(* IEC 61131-3 sources: Caravan/Archiv/12-04-19/Stations/MachineControl/MachineControl/Class/SafetyManager (part 2) *)

	state := READY;

//=================================================================================================
#ifdef VM_CLASS_TIME_MEASUREMENT
	StopTimeMeasurement(VARANTIME_CY);
#endif
//=================================================================================================

END_FUNCTION

FUNCTION SafetyManager::AddModule
	VAR_INPUT
		pPara 	: ^CmdStruct;
	END_VAR
	VAR_OUTPUT
		retcode 	: BOOL;
	END_VAR
  VAR
  	ModuleType : t_e_ModuleType;
  END_VAR

  retcode := FALSE;

  ModuleType := pPara^.aPara[0]$t_e_ModuleType;

  // we differ between real safety components and managing components
  case ModuleType of
    _CSCP01x,
    _CSDI16x,
    _CSTO08x,
    _SCP010,
    _SCP011,
    _SCP111,
    _MS011,
    _MS012,
    _SDD1300,
    _SDD1400,
    _SDD1500,
    _SDD1600:
        retcode := AddSafetyModule(ModuleType, pPara^.aPara[1]$pVirtualBase);

        if IsFSoEModule(ModuleType) then
          // allocate memory for the temporary cyclic send buffer
          sUdpVars.pTempSendBufferCy$pVoid := To_StdLib.Malloc(size:=sizeof(t_UdpPacket));

          if sUdpVars.pTempSendBufferCy then
            _memset(dest:=sUdpVars.pTempSendBufferCy, usByte:=0, cntr:=sizeof(t_UdpPacket));
          else
            SetError(bError:=TRUE, ErrorMessage:=_NO_MEMORY_SENDBUFFER_UDP_ERROR, dError:=0);
            LogError("@ZZZZ (SafetyManager::AddModule) Failed to allocate memory for udp send buffer");
          end_if;

          // allocate memory for the temporary irq send buffer
          sUdpVars.pTempSendBufferIRQ$pVoid := To_StdLib.Malloc(size:=sizeof(t_UdpPacket));

          if sUdpVars.pTempSendBufferIRQ then
            _memset(dest:=sUdpVars.pTempSendBufferIRQ, usByte:=0, cntr:=sizeof(t_UdpPacket));
          else
            SetError(bError:=TRUE, ErrorMessage:=_NO_MEMORY_SENDBUFFER_UDP_ERROR, dError:=0);
            LogError("@ZZZZ (SafetyManager::AddModule) Failed to allocate memory for udp send buffer");
          end_if;

          sUdpVars.paConnectionsToProducers$pVoid := To_StdLib.Malloc(size:=sizeof(t_aUdpConnections));

          if sUdpVars.paConnectionsToProducers then
            _memset(dest:=sUdpVars.paConnectionsToProducers, usByte:=0, cntr:=sizeof(t_aUdpConnections));
          else
            SetError(bError:=TRUE, ErrorMessage:=_NO_MEMORY_CONNECTION_BUFFER_UDP_ERROR, dError:=0);
            LogError("@ZZZZ (SafetyManager::AddModule) Failed to allocate memory for udp receive buffer");
          end_if;

          sUdpVars.paConnectionsToConsumers$pVoid := To_StdLib.Malloc(size:=sizeof(t_aUdpConnections));

          if sUdpVars.paConnectionsToConsumers then
            _memset(dest:=sUdpVars.paConnectionsToConsumers, usByte:=0, cntr:=sizeof(t_aUdpConnections));
          else
            SetError(bError:=TRUE, ErrorMessage:=_NO_MEMORY_CONNECTION_BUFFER_UDP_ERROR, dError:=0);
            LogError("@ZZZZ (SafetyManager::AddModule) Failed to allocate memory for udp receive buffer");
          end_if;
        end_if;

    _VBC021Master,
    _VBC021Slave, // (is limited to 1 per system, because the system can't sync to different systems at the same time)
    _VMC052,
    _VaranManager4VMC, // VaranManager (VMC052 counterpart is also limited to 1 per system, because the system can't sync to different systems at the same time)
    _GenericTimeSyncMaster,
    _GenericTimeSyncSlave:
        retcode := AddManagingModule(ModuleType, pPara^.aPara[1]$pVirtualBase, pPara^.aPara[2]$^USINT);
  else
    // invalid module type
    ClassState := -7;
    LogError("@ZZZZ (SafetyManager::AddModule) Invalid ModuleType");
  end_case;

  if retcode then
    LoginCnt += 1;
  end_if;

END_FUNCTION

FUNCTION SafetyManager::AddSafetyModule
	VAR_INPUT
		ModuleType 	: t_e_ModuleType;
		pThis 	: pVirtualBase;
	END_VAR
	VAR_OUTPUT
		retcode 	: BOOL;
	END_VAR
  VAR
  	pHelpSafety : ^t_SafetyComponent;
  END_VAR

  if pFirstSafetyComponent = NIL then
    pFirstSafetyComponent$pVoid := To_StdLib.Malloc(size:=sizeof(t_SafetyComponent));
    pHelpSafety := pFirstSafetyComponent;
  else
    pHelpSafety := pFirstSafetyComponent;
    while pHelpSafety^.pNext <> NIL do
      pHelpSafety := pHelpSafety^.pNext;
    end_while;
    pHelpSafety^.pNext$pVoid := To_StdLib.Malloc(size:=sizeof(t_SafetyComponent));
    pHelpSafety := pHelpSafety^.pNext;
  end_if;

  if pHelpSafety <> NIL then
    _memset(dest:=pHelpSafety, usByte:=0, cntr:=sizeof(t_SafetyComponent));
    pHelpSafety^.ModuleType   := ModuleType;
    pHelpSafety^.pThis        := pThis;

//    pHelpSafety^.pNext        := NIL;  // not necessary because of memset

    case ModuleType of
//**********************************************************************************************************************************************************
      _CSCP01x,
      _SCP010,
      _SCP011,
      _SCP111,
      _SDD1300,
      _SDD1400,
      _SDD1500,
      _SDD1600:
        LocalCPUNo += 1;

//**********************************************************************************************************************************************************
      _CSDI16x,
      _MS011,
      _MS012:
        pHelpSafety^.InfoBits.OnlyInputs := TRUE;
//**********************************************************************************************************************************************************
    end_case;

    us_SafetyModuleNo += 1;

    retcode := TRUE;
  else
    ClassState := -1;

    retcode := FALSE;
  end_if;

END_FUNCTION

FUNCTION SafetyManager::AddManagingModule
	VAR_INPUT
		ModuleType 	: t_e_ModuleType;
		pThis 	: pVirtualBase;
		pObjectPath 	: ^USINT;
	END_VAR
	VAR_OUTPUT
		retcode 	: BOOL;
	END_VAR
  VAR
  	pHelpManaging : ^t_ManagingComponent;
    pMyPath : ^USINT;
  END_VAR

  if pFirstManagingInterfaceComponent = NIL then
    pFirstManagingInterfaceComponent$pVoid := To_StdLib.Malloc(size:=sizeof(t_ManagingComponent));
    pHelpManaging := pFirstManagingInterfaceComponent;
  else
    pHelpManaging := pFirstManagingInterfaceComponent;
    while pHelpManaging^.pNext <> NIL do
      pHelpManaging := pHelpManaging^.pNext;
    end_while;
    pHelpManaging^.pNext$pVoid := To_StdLib.Malloc(size:=sizeof(t_ManagingComponent));
    pHelpManaging := pHelpManaging^.pNext;
  end_if;

  if pHelpManaging <> NIL then
    _memset(dest:=pHelpManaging, usByte:=0, cntr:=sizeof(t_ManagingComponent));
    pHelpManaging^.ModuleType     := ModuleType;
    pHelpManaging^.pThis          := pThis;
    pHelpManaging^.DomainNr       := 16#FF;

    if pObjectPath then
      pMyPath$^void := To_StdLib.Malloc(size:=pObjectPath^ + 2);

      // convert 1 byte length info into 2 byte length info
      if pMyPath then
        pMyPath^$UINT := pObjectPath^$USINT;
        To_StdLib.MemCpy(dest:=pMyPath + 2, source:=pObjectPath + 1, size:=pObjectPath^);
      end_if;
    end_if;

    pHelpManaging^.pModulePath := pMyPath;

  //pHelpManaging^.pNext          := NIL;  // not necessary because of memset

    retcode := TRUE;
  else
    ClassState := -1;

    retcode := FALSE;
  end_if;

END_FUNCTION

FUNCTION SafetyManager::AddSafetyNbr
	VAR_INPUT
		pThis 	: pVirtualBase;
		ud_SafetyNbr 	: UDINT;
		FirmwareVersion 	: HDINT;
		FPGAVersion 	: HSINT;
		PathLen 	: USINT;
		pPath 	: ^USINT;
	END_VAR
	VAR_OUTPUT
		retcode 	: BOOL;
	END_VAR
  VAR
  	pHelpSafety : ^t_SafetyComponent;
  END_VAR

  retcode := FALSE;

  if pFirstSafetyComponent then
    pHelpSafety := pFirstSafetyComponent;
    while pHelpSafety do
      if pHelpSafety^.pThis = pThis then
        pHelpSafety^.SafetyNbr    := ud_SafetyNbr;
        pHelpSafety^.FW_Version   := FirmwareVersion;
        pHelpSafety^.FPGA_Version := FPGAVersion;
        pHelpSafety^.PathLen      := PathLen;
        pHelpSafety^.pPath        := pPath;

        // look for local safety CPU
        if b_CheckSafetyTopology then
          if (PathLen > 2) & (((pPath+2)^ = HWT_ESCAPE_CDIAS) | ((pPath+2)^ = HWT_ESCAPE_SDIAS)) then
            b_CheckSafetyTopology := FALSE; // Safety-CPU is local -> no problem
          end_if;
        end_if;

        retcode := TRUE;
        return;
      end_if;

      pHelpSafety := pHelpSafety^.pNext;
    end_while;
  end_if;

END_FUNCTION

FUNCTION SafetyManager::GetModuleTypeNo
	VAR_INPUT
		ModuleType 	: t_e_ModuleType;
	END_VAR
	VAR_OUTPUT
		ModuleNo 	: DINT;
	END_VAR
  VAR
  	pHelpSafety   : ^t_SafetyComponent;
    pHelpManaging : ^t_ManagingComponent;
  END_VAR

  ModuleNo := 0;

  if pFirstSafetyComponent then
    pHelpSafety := pFirstSafetyComponent;
    while pHelpSafety do
      if pHelpSafety^.ModuleType = ModuleType then
        ModuleNo += 1;
      end_if;

      pHelpSafety := pHelpSafety^.pNext;
    end_while;
  end_if;

  if pFirstManagingInterfaceComponent then
    pHelpManaging := pFirstManagingInterfaceComponent;
    while pHelpManaging do
      if pHelpManaging^.ModuleType = ModuleType then
        ModuleNo += 1;
      end_if;

      pHelpManaging := pHelpManaging^.pNext;
    end_while;
  end_if;

END_FUNCTION

FUNCTION SafetyManager::NewTimeSyncPossible
	VAR_OUTPUT
		retcode 	: BOOL;
	END_VAR
  VAR
  	pHelpSafety   : ^t_SafetyComponent;
  END_VAR

  // if there is FSoE in the project => no timesync
  if b_GotFSoEModules then
    retcode := FALSE;
    return;
  end_if;

  // default is: we can => check if there is any module with too old firmware or fpga
  retcode := TRUE;

  if pFirstSafetyComponent then
    pHelpSafety := pFirstSafetyComponent;
    while pHelpSafety do

      // check all modules for correct versions
      if ((pHelpSafety^.ModuleType = _CSCP01x) & (   (pHelpSafety^.FPGA_Version    < 16#14)     // if its a CSCP and the FPGA Version is lower than 1.4
                                                   | (pHelpSafety^.FW_Version$UINT < 100)) &    // or the firmware version is lower than 100
                                                      pHelpSafety^.SafetyNbr)                   // only if there is a safety number available (maybe the module is optional and not available)
      |  (pHelpSafety^.NewConfigType = ConfigState_Old) then                                    // or the module has an old config type

        retcode := FALSE;
      end_if;

      pHelpSafety := pHelpSafety^.pNext;
    end_while;
  end_if;

END_FUNCTION

FUNCTION SafetyManager::SetNewSyncMode
	VAR_INPUT
		b_NewMode 	: BOOL;
	END_VAR
  VAR
		MyPara 	  : CmdStruct;
		MyResult	: results;
  END_VAR

  b_NewSyncMode := b_NewMode;

  MyPara.uiCmd := CMD_SM_SET_NEW_SYNC_MODE;
  MyPara.aPara[0] := b_NewSyncMode;
  TellAllSafetyModules(#MyPara, #MyResult);

END_FUNCTION

FUNCTION SafetyManager::TellAllSafetyModules
	VAR_INPUT
		pPara 	: ^CmdStruct;
		pResult 	: ^results;
	END_VAR
  VAR
  	pHelpSafety : ^t_SafetyComponent;
  END_VAR

  if pFirstSafetyComponent then
    pHelpSafety := pFirstSafetyComponent;
    while pHelpSafety do
      // call the newinst with the given parameters
      pHelpSafety^.pThis^.NewInst(pPara, pResult);

      pHelpSafety := pHelpSafety^.pNext;
    end_while;
  end_if;

END_FUNCTION

FUNCTION SafetyManager::StartTimeSync

  if pFirstTimeSyncElement then
    pActTimeSyncElement := pFirstTimeSyncElement;

    // send the token to the right module
    GiveTokenToNextModule();

    // remember the start time for calculating the time of a complete synchronisation
    TimeSyncCycleStart := ops.tAbsolute;
  end_if;

END_FUNCTION

FUNCTION SafetyManager::NextTimeSyncModule

  pActTimeSyncElement := pActTimeSyncElement^.pNext;

  // must be done after selecting the new element
  if GiveTokenToNextModule() then
    // we're finished with our synchronisation cycle and just started a new one (must be done after selecting the new element)
    if IsTimeSyncMaster then
      SyncDuration := ops.tAbsolute - TimeSyncCycleStart;
      if SyncDuration > MaxSyncDuration then
        MaxSyncDuration := SyncDuration;
      end_if;
      if SyncDuration < MinSyncDuration then
        MinSyncDuration := SyncDuration;
      end_if;

      // if a cycle has been finished => reset the timeout counter
      SyncTimeoutCounter := 0;

      // remember the start time for calculating the time of a complete synchronisation
      TimeSyncCycleStart := ops.tAbsolute;
    end_if;
  end_if;

END_FUNCTION

FUNCTION SafetyManager::GiveTokenToNextModule
	VAR_OUTPUT
		RestartCycle 	: BOOL;
	END_VAR
  VAR
		MyPara 	  : CmdStruct;
		MyResult	: results;
    pTemp : ^t_TimeSyncElement;
  END_VAR

  if pActTimeSyncElement = pFirstTimeSyncElement then
    RestartCycle := TRUE;
  else
    RestartCycle := FALSE;
  end_if;

  // check if we have to skip something (missing optional modules)
  if TimeSyncModuleAvailable(pActTimeSyncElement) = FALSE then
    // save the actual position
    pTemp := pActTimeSyncElement;

    // if it's a missing optional module
    while (TimeSyncModuleAvailable(pActTimeSyncElement) = FALSE) do
      // skip it
      pActTimeSyncElement := pActTimeSyncElement^.pNext;

      // if we jumped on the first, we have to restart the cycle (time measurement and timeout surveillance)
      if pActTimeSyncElement = pFirstTimeSyncElement then
        RestartCycle := TRUE;
      end_if;

      // if we're at the start of the rotation => stop rotating and print error message
      if pActTimeSyncElement = pTemp then
        bd_LogRtMessagesInCy.TooManyOptionalMissing := TRUE;
        ClassState := -12;
        exit;
      end_if;
    end_while;
  end_if;

  // check if we have to skip something
  if pActTimeSyncElement^.InfoBits.IsInterfaceDomain then
    // save the actual position
    pTemp := pActTimeSyncElement;

    // if it's an interface managing module and it's not synchron, skip it (there has to be also a Safety CPU in the system, therefore we don't ask for it
    while pActTimeSyncElement^.InfoBits.IsInterfaceDomain & (pActTimeSyncElement^.pManaging^.InfoBits.IsSynchron = FALSE) do
      // skip it
      pActTimeSyncElement := pActTimeSyncElement^.pNext;

      // if we jumped on the first, we have to restart the cycle (time measurement and timeout surveillance)
      if pActTimeSyncElement = pFirstTimeSyncElement then
        RestartCycle := TRUE;
      end_if;

      // if we're at the start of the rotation => stop rotating and print error message
      if pActTimeSyncElement = pTemp then
        bd_LogRtMessagesInCy.InvalidIFConfiguration := TRUE;
        ClassState := -12;
        exit;
      end_if;
    end_while;
  end_if;

  if pActTimeSyncElement^.InfoBits.IsConnectionToMaster then
    // don't check for sync timeout if we're not the master
    b_CheckTimeSyncTimeout := FALSE;
  else
    b_CheckTimeSyncTimeout := TRUE;
  end_if;

  // if it's a managing module and not the connection to the master, we give the token to a slave => remember it
  if pActTimeSyncElement^.InfoBits.IsManagingModule & (pActTimeSyncElement^.InfoBits.IsConnectionToMaster = FALSE) then
    b_SlaveSyncActive := TRUE;
  end_if;

  // tell the next module, to start the time synchronisation
  MyPara.uiCmd := CMD_SM_START_TIME_SYNC;
  pActTimeSyncElement^.pThis^.NewInst(#MyPara, #MyResult);

  LastTimeSyncThis := pActTimeSyncElement^.pThis;
  TimeSyncTimeStamp := ops.tAbsolute;

END_FUNCTION

FUNCTION SafetyManager::TellAllInterfaceManagingModules
	VAR_INPUT
		pPara 	: ^CmdStruct;
		pResult 	: ^results;
		OverrideSync 	: BOOL;(* := FALSE *)
	END_VAR
  VAR
  	pHelpManaging : ^t_ManagingComponent;
  END_VAR

  if pFirstManagingInterfaceComponent then
    pHelpManaging := pFirstManagingInterfaceComponent;
    while pHelpManaging do
      // call the newinst with the given parameters
      if pHelpManaging^.InfoBits.IsSynchron | OverrideSync then
        pHelpManaging^.pThis^.NewInst(pPara, pResult);
      end_if;

      pHelpManaging := pHelpManaging^.pNext;
    end_while;
  end_if;

END_FUNCTION

FUNCTION SafetyManager::SafetyManager
	VAR_OUTPUT
		ret_code 	: ConfStates;
	END_VAR
  VAR
    sd_retval : DINT;
  END_VAR

  //get interface for hardwaretree functions
  if ( OS_CILGET(INTERFACE_HARDWARETREE, #pHardwareTree)) then
    pHardwareTree := NIL;

    // logging can be used here already because the constructor of the base has been called before to initialize the log-interface-pointer
    LogError("@ZZZZ (SafetyManager::SafetyManager) Hardwaretree-Interface not found. A newer OS is required for Safety-Modules");
  end_if;

  pTempMemCy := To_StdLib.Malloc(size:=SIZE_TEMP_MEMORY);
  if pTempMemCy then
    ud_SizeTempMemCy := SIZE_TEMP_MEMORY;
  else
    LogError("@ZZZZ (SafetyManager::SafetyManager) Allocate temporary Memory failed");
  end_if;

  b_QuitErrorAvailable := FALSE;

  sd_retval := OS_CILGet(INTERFACE_SAFETY_DLL, #pSafetyDll)$DINT;

  if sd_retval then
    // normal case => no dll available
//    LogValue("@ZZZZ (SafetyManager::SafetyManager) Failed to get interface to safety DLL with ErrorCode 0x{0}", Value:=sd_retval$UDINT);
  elsif pSafetyDll^.version >= 5 then
//    LogValue("@ZZZZ (SafetyManager::SafetyManager) Safety DLL with Version 0x{0} loaded. QuitError via Application available!", Value:=pSafetyDll^.version);

    b_QuitErrorAvailable := TRUE;
  end_if;

  // as long there is no Safety-CPU on local CDIAS or SDIAS, we need to check for "unalowed" safety communication over VARAN.
  b_CheckSafetyTopology := TRUE;
  OS_CILGet( INTERFACE_VARANMANAGER, #pVaran );

	ret_code := C_OK;

END_FUNCTION

FUNCTION SafetyManager::AllManagingNodesSynchron
	VAR_OUTPUT
		AllReady 	: BOOL;
	END_VAR
  VAR
  	pHelpManaging : ^t_ManagingComponent;
		MyPara 	  : CmdStruct;
		MyResult	: results;
  END_VAR

  AllReady := TRUE;

  // check if any of the managing interface modules is not synchron
  if pFirstManagingInterfaceComponent then
    MyPara.uiCmd := CMD_SM_SYNC_CHECK;

    pHelpManaging := pFirstManagingInterfaceComponent;
    while pHelpManaging do
      // if any managing component isn't synchron => stop searching
      if pHelpManaging^.pThis^.NewInst(#MyPara, #MyResult) = ERROR then
        if (pHelpManaging^.InfoBits.IsOptional = TRUE) then
          if ((SafetyDomainTimeout & ((ops.tAbsolute - SynchroTimeout) > SafetyDomainTimeout))) then
            // we give up waiting => timeout exceeded
            b_SyncTimeoutExceeded := TRUE;
            // if it's the last managing module, then it's our connection to the master module
            if (IsTimeSyncMaster = 0) & pHelpManaging^.InfoBits.IsConnectionToMaster then
              // we have to be our own master now
              IsTimeSyncMaster := 1;
            end_if;
          else
            AllReady := FALSE;
          end_if;
        else
          AllReady := FALSE;
        end_if;

        // return; don't give up here => we have to check it for all domains, this one may be an optional interface frame domain
        pHelpManaging^.InfoBits.IsSynchron := FALSE;
      else
        pHelpManaging^.InfoBits.IsSynchron := TRUE;
      end_if;

      pHelpManaging := pHelpManaging^.pNext;
    end_while;
  end_if;

END_FUNCTION

FUNCTION SafetyManager::GetMasterConnection
  VAR_OUTPUT
    pMasterConn : ^t_ManagingComponent;
  END_VAR
  VAR
    pHelpManaging : ^t_ManagingComponent;
  END_VAR

  pMasterConn := NIL;

  if pFirstManagingInterfaceComponent then
    pHelpManaging := pFirstManagingInterfaceComponent;
    while pHelpManaging do
      if (pHelpManaging^.ModuleType = _VBC021Slave) | (pHelpManaging^.ModuleType = _VaranManager4VMC) | (pHelpManaging^.ModuleType = _GenericTimeSyncSlave) then
        pMasterConn := pHelpManaging;
        pMasterConn^.InfoBits.IsConnectionToMaster := TRUE;
        // if it's not the last in the list => we have to put it in the last place for easier timesync handling (last managing module to handle is the connection back to the master)
        if pMasterConn^.pNext then
          // if it's the first one
          if pMasterConn = pFirstManagingInterfaceComponent then
            pHelpManaging := pFirstManagingInterfaceComponent;
            while pHelpManaging^.pNext do
              pHelpManaging := pHelpManaging^.pNext;
            end_while;
            pFirstManagingInterfaceComponent := pFirstManagingInterfaceComponent^.pNext;
            pHelpManaging^.pNext := pMasterConn;
            pMasterConn^.pNext := NIL;
          else
            // if it's one in the middle
            pHelpManaging := pFirstManagingInterfaceComponent;
            while pHelpManaging^.pNext do
              if pHelpManaging^.pNext = pMasterConn then
                pHelpManaging^.pNext := pMasterConn^.pNext;
              end_if;

              pHelpManaging := pHelpManaging^.pNext;
            end_while;
            pHelpManaging^.pNext := pMasterConn;
            pMasterConn^.pNext := NIL;
          end_if;
        end_if;
        return;
      end_if;

      pHelpManaging := pHelpManaging^.pNext;
    end_while;
  end_if;

END_FUNCTION

FUNCTION SafetyManager::AddConfiguration
	VAR_INPUT
		Length 	: UINT;
		pData 	: ^void;
		IsFSoEConfig 	: BOOL;
	END_VAR
	VAR_OUTPUT
		retcode 	: DINT;
	END_VAR
  VAR
    pHelpCfg          : ^t_CfgListElem;
    pHelpModule       : ^t_ModuleListElem;
    pHelpPdo          : ^t_PdoListElem;
    pHelpSlave        : ^t_SlaveListElem;
    pHelpConnection   : ^t_FSoEConnectionDetails;
    pDataHelp         : ^void;
    i                 : UDINT;
    TmpPathLen        : UINT;
    TempCfgNo         : USINT;
    TempConnectionNo  : UINT;
  END_VAR

(*
    Memory structure:
      4 Byte: SafetyNumber of CPU (is already there from initialisation in CSCP011_IM::InitSafeModule)
      1 Byte: Number of module configurations which are following
      for every module configuration (first is always the CPU itself)
        1 Byte: Info
        4 Byte: Interface Frame Source SafetyNumber (0 if it is no source for interface frames)
        4 Byte: Interface Frame CRC
        1 Byte: Number of destination inferface frame CRCs
        x Byte: Destination interface frame CRCs (number * sizeof(HDINT)
        2 Byte: Length of hardware path
        x Byte (depending on length in the 2 byte before): Hardwarepath
        2 Byte: Length of compressed hardware path
        x Byte (depending on length in the 2 byte before): Compressed Hardwarepath
        1 Byte: PDO out length for this module
      1 Byte: Number of pdo configurations which are following
      for every PDO configuration
        1 Byte: PDO length
        1 Byte: Interface frame info
        4 Byte: Interface CRC
        2 Byte: Length of source hardware path
        x Byte (depending on length in the 2 byte before): Hardwarepath of source
        2 Byte: Length of destination hardware path
        x Byte (depending on length in the 2 byte before): Hardwarepath of destination
      1 Byte: Number of slave configurations which are following
      for every slave configuration
        1 Byte: Info
        4 Byte: InterfaceCRC
        2 Byte: Length of hardware path
        x Byte (depending on length in the 2 byte before): Hardwarepath
        2 Byte: Length of compressed hardware path
        x Byte (depending on length in the 2 byte before): Compressed Hardwarepath

      if IsFSoEConfig = TRUE
      2 Byte: Number of connection infos which are following
      for every FSoE connection info
        2 Byte: ConnectionID
        1 Byte: ConnectionState
        1 Byte: Flags // Actually, type is 4 bytes in size but for compatibility reasons it is still used as 1 byte. As a result, bits 9-32 are currently not used.
        4 Byte: Master safety number

only if feature available:
        2 Byte: Transmission time in ms

        2 Byte: Offset where to read from master
        2 Byte: Size of data to read from master (and write to slave)
        2 Byte: Offset where to write to master
        2 Byte: Size of data to write to master (and read from slave)
        2 Byte: SlaveAddress
        2 Byte: Length of slave hardware path
        x Byte (depending on length in the 2 byte before): Slave hardware path
        2 Byte: Length of compressed slave hardware path
        x Byte (depending on length in the 2 byte before): Compressed slave hardware path
        2 Byte: Offset where to read from slave
        2 Byte: Offset where to write to slave

*)

  // check if the configuration is valid (pData <> NIL) & (Length must be at least 4 byte for SafetyNbr + 1 byte module cfg number + 1 byte pdo cfg number + 1 byte slave cfc number)
  if pData & (Length >= 7)  then

    retcode := 0;

    // first we have to allocate some memory for the configuration
    if pConfigs = NIL then
      pConfigs$pVoid := To_StdLib.Malloc(size:=sizeof(t_CfgListElem));
      pHelpCfg := pConfigs;
    else
      pHelpCfg := pConfigs;
      while pHelpCfg^.pNext <> NIL do
        //if searched path is found, we already got this module in our list
        if pHelpCfg^.SafetyNbr = pData^$HDINT then
          // already in buffer => leave function
          return;
        else
          pHelpCfg := pHelpCfg^.pNext;
        end_if;
      end_while;

      //if searched path is found, we already got this module in our list
      if pHelpCfg^.SafetyNbr = pData^$HDINT then
        // already in buffer => leave function
        return;
      end_if;

      pHelpCfg^.pNext$pvoid := To_StdLib.Malloc(size:=sizeof(t_CfgListElem));
      pHelpCfg := pHelpCfg^.pNext;
    end_if;

    // if we have memory for the configuration => we add the data to the new element
    if pHelpCfg <> NIL then
      pDataHelp := pData;

      // set the next pointer to NIL
      pHelpCfg^.pNext := NIL;

      // safety number of the safety cpu
      pHelpCfg^.SafetyNbr := pDataHelp^$HDINT;
      pDataHelp += sizeof(HDINT);

      // number of module configurations which follow now
      TempCfgNo := pDataHelp^$USINT;
      pDataHelp += sizeof(USINT);

      pHelpCfg^.pFirstModuleCfg := NIL;

      // module configurations
      if TempCfgNo then
        for i := 0 to (TempCfgNo-1) do
          if pHelpCfg^.pFirstModuleCfg = NIL then
            pHelpCfg^.pFirstModuleCfg$pVoid := To_StdLib.Malloc(size:=sizeof(t_ModuleListElem));
            pHelpModule := pHelpCfg^.pFirstModuleCfg;
          else
            pHelpModule^.pNext$pvoid := To_StdLib.Malloc(size:=sizeof(t_ModuleListElem));
            pHelpModule := pHelpModule^.pNext;
          end_if;

          if pHelpModule then
            // initialize the pointers with NIL in case one of the mallocs fails
            pHelpModule^.ModuleInfo.pDestCRCs   := NIL;
            pHelpModule^.ModuleInfo.pPath       := NIL;
            pHelpModule^.ModuleInfo.pCompPath   := NIL;
            pHelpModule^.pNext                  := NIL;

            // info
            pHelpModule^.ModuleInfo.Info := pDataHelp^$BSINT;
            pDataHelp += sizeof(BSINT);

            // safety number of interface frame source
            pHelpModule^.ModuleInfo.SafetyNbr := pDataHelp^$HDINT;
            pDataHelp += sizeof(HDINT);

            // interface CRC of interface frame
            pHelpModule^.ModuleInfo.InterfaceCRC := pDataHelp^$HDINT;
            pDataHelp += sizeof(HDINT);

            if pHelpModule^.ModuleInfo.InterfaceCRC then
              // someone might connect to us via udp because we supply an interface frame
              sUdpVars.UdpInit.ProvidesIF := TRUE;
            end_if;

            // interface frame destination CRCs
            if pHelpModule^.ModuleInfo.Info.IsInterfaceDest then
              // number of CRCs
              TmpPathLen := pDataHelp^$USINT; // save some time with this local variable
              pHelpModule^.ModuleInfo.DestCRCNo := TmpPathLen$USINT;
              pDataHelp += sizeof(USINT);

              // allocate memory for the module path
              pHelpModule^.ModuleInfo.pDestCRCs$pVoid := To_StdLib.Malloc(size:=TmpPathLen * sizeof(HDINT));
              if pHelpModule^.ModuleInfo.pDestCRCs = NIL then
                ClassState := -1;
                retcode := -2;
                return;
              end_if;

              // save CRCs
              _memcpy(ptr1:=pHelpModule^.ModuleInfo.pDestCRCs, ptr2:=pDataHelp, cntr:=TmpPathLen * sizeof(HDINT));
              pDataHelp += TmpPathLen * sizeof(HDINT);
            else
              pHelpModule^.ModuleInfo.DestCRCNo := 0;
              pHelpModule^.ModuleInfo.pDestCRCs := NIL;
            end_if;

            // length of hardwarepath
            TmpPathLen := pDataHelp^$UINT; // save some time with this local variable
            pHelpModule^.ModuleInfo.PathLen := TmpPathLen;
            pDataHelp += sizeof(UINT);

            // allocate memory for the module path
            pHelpModule^.ModuleInfo.pPath$pVoid := To_StdLib.Malloc(size:=TmpPathLen);
            if pHelpModule^.ModuleInfo.pPath = NIL then
              ClassState := -1;
              retcode := -2;
              return;
            end_if;

            // save hardwarepath
            _memcpy(ptr1:=pHelpModule^.ModuleInfo.pPath, ptr2:=pDataHelp, cntr:=TmpPathLen);
            pDataHelp += TmpPathLen;

            // length of hardwarepath
            TmpPathLen := pDataHelp^$UINT; // save some time with this local variable
            pHelpModule^.ModuleInfo.CompPathLen := TmpPathLen;
            pDataHelp += sizeof(UINT);

            // allocate memory for the module path
            pHelpModule^.ModuleInfo.pCompPath$pVoid := To_StdLib.Malloc(size:=TmpPathLen);
            if pHelpModule^.ModuleInfo.pCompPath = NIL then
              ClassState := -1;
              retcode := -2;
              return;
            end_if;

            // save compressed hardwarepath
            _memcpy(ptr1:=pHelpModule^.ModuleInfo.pCompPath, ptr2:=pDataHelp, cntr:=TmpPathLen);
            pDataHelp += TmpPathLen;

            // PDO out length for this module (to assign the length to the pdo configurations)
            pHelpModule^.ModuleInfo.PdoOutLen := pDataHelp^$USINT;
            pDataHelp += sizeof(USINT);
          else
            ClassState := -1;
            retcode := -2;
            return;
          end_if;
        end_for;
      end_if;

      // number of Pdo configurations which follow now
      TempCfgNo := pDataHelp^$USINT;
      pDataHelp += sizeof(USINT);

      pHelpCfg^.pFirstPdoCfg := NIL;

      // Pdo configurations
      if TempCfgNo then
        for i := 0 to (TempCfgNo-1) do
          if pHelpCfg^.pFirstPdoCfg = NIL then
            pHelpCfg^.pFirstPdoCfg$pVoid := To_StdLib.Malloc(size:=sizeof(t_PdoListElem));
            pHelpPdo := pHelpCfg^.pFirstPdoCfg;
          else
            pHelpPdo^.pNext$pvoid := To_StdLib.Malloc(size:=sizeof(t_PdoListElem));
            pHelpPdo := pHelpPdo^.pNext;
          end_if;

          if pHelpPdo then
            // initialize the pointers with NIL in case one of the mallocs fails
            pHelpPdo^.PdoInfo.pSourcePath     := NIL;
            pHelpPdo^.PdoInfo.pDestPath       := NIL;
            pHelpPdo^.pNext                   := NIL;

            // pdo length
            pHelpPdo^.PdoInfo.PdoLen := pDataHelp^$USINT;
            pDataHelp += sizeof(USINT);

            // is it an interface pdo?
            pHelpPdo^.PdoInfo.Info := pDataHelp^$BSINT;
            pDataHelp += sizeof(BSINT);

            // if it is an interface frame, we have to copy the CRC too
            if pHelpPdo^.PdoInfo.Info.IsInterfacePDO then
              // interface CRC
              pHelpPdo^.PdoInfo.InterfaceCRC := pDataHelp^$HDINT;
            else
              pHelpPdo^.PdoInfo.InterfaceCRC := 0;
            end_if;
            pDataHelp += sizeof(HDINT);

            // length of source hardwarepath
            TmpPathLen := pDataHelp^$UINT; // save some time with this local variable
            pHelpPdo^.PdoInfo.SourcePathLen := TmpPathLen;
            pDataHelp += sizeof(UINT);

            // allocate memory for the source module path
            pHelpPdo^.PdoInfo.pSourcePath$pVoid := To_StdLib.Malloc(size:=TmpPathLen);
            if pHelpPdo^.PdoInfo.pSourcePath = NIL then
              ClassState := -1;
              retcode := -2;
              return;
            end_if;

            // save source hardwarepath
            _memcpy(ptr1:=pHelpPdo^.PdoInfo.pSourcePath, ptr2:=pDataHelp, cntr:=TmpPathLen);
            pDataHelp += TmpPathLen;

            // check for an IP Address
            if pHelpPdo^.PdoInfo.Info.SrcPathIsCompressed & (pHelpPdo^.PdoInfo.pSourcePath^$USINT = INTERFACE_IP_MODE) then
              // add the connection (we're consumer and we got the IP address of the producer)
              AddUdpConnection(IP:=(pHelpPdo^.PdoInfo.pSourcePath$^HDINT + 5)^, IFCRC:=(pHelpPdo^.PdoInfo.pSourcePath$^HDINT + 1)^, SafetyNumber:=pHelpCfg^.SafetyNbr, ProducerList:=TRUE);
            end_if;

            // length of destination hardwarepath
            TmpPathLen := pDataHelp^$UINT; // save some time with this local variable
            pHelpPdo^.PdoInfo.DestPathLen := TmpPathLen;
            pDataHelp += sizeof(UINT);

            // allocate memory for the destination module path
            pHelpPdo^.PdoInfo.pDestPath$pVoid := To_StdLib.Malloc(size:=TmpPathLen);
            if pHelpPdo^.PdoInfo.pDestPath = NIL then
              ClassState := -1;
              retcode := -2;
              return;
            end_if;

            // save destination hardwarepath
            _memcpy(ptr1:=pHelpPdo^.PdoInfo.pDestPath, ptr2:=pDataHelp, cntr:=TmpPathLen);
            pDataHelp += TmpPathLen;

            // check if a prior configuration also added this PDO (possible if a CSTO gets PDOs from 2 CSCPs)
            if DoublePDOEntry(pHelpPdo^.PdoInfo, pHelpCfg) then
              // use ID 255 (as kind of invalid) and mark the PDO as double entry (will not be distributed then)
              pHelpPdo^.PdoInfo.PDO_ID := 255;
              pHelpPdo^.PdoInfo.Info.DoublePDOEntry := TRUE;
            else
              // now we give it a priority and increase the number for the next pdo
              pHelpPdo^.PdoInfo.PDO_ID := ActPDO_ID;
              ActPDO_ID += 1;
            end_if;

          else
            ClassState := -1;
            retcode := -2;
            return;
          end_if;
        end_for;
      end_if;

      // number of slave configurations which follow now
      TempCfgNo := pDataHelp^$USINT;
      pDataHelp += sizeof(USINT);

      pHelpCfg^.pFirstSlaveCfg:= NIL;

      // slave configurations
      if TempCfgNo then
        for i := 0 to (TempCfgNo-1) do
          if pHelpCfg^.pFirstSlaveCfg = NIL then
            pHelpCfg^.pFirstSlaveCfg$pVoid := To_StdLib.Malloc(size:=sizeof(t_SlaveListElem));
            pHelpSlave := pHelpCfg^.pFirstSlaveCfg;
          else
            pHelpSlave^.pNext$pvoid := To_StdLib.Malloc(size:=sizeof(t_SlaveListElem));
            pHelpSlave := pHelpSlave^.pNext;
          end_if;

          if pHelpSlave then
            // initialize the pointers with NIL in case one of the mallocs fails
            pHelpSlave^.SlaveInfo.pPath     := NIL;
            pHelpSlave^.SlaveInfo.pCompPath := NIL;
            pHelpSlave^.pNext               := NIL;

            // info
            pHelpSlave^.SlaveInfo.Info := pDataHelp^$BSINT;
            pDataHelp += sizeof(BSINT);

            // InterfaceCRC
            pHelpSlave^.SlaveInfo.InterfaceCRC := pDataHelp^$HDINT;
            pDataHelp += sizeof(HDINT);

            // length of hardwarepath
            TmpPathLen := pDataHelp^$UINT; // save some time with this local variable
            pHelpSlave^.SlaveInfo.PathLen := TmpPathLen;
            pDataHelp += sizeof(UINT);

            // allocate memory for the module path
            pHelpSlave^.SlaveInfo.pPath$pVoid := To_StdLib.Malloc(size:=TmpPathLen);
            if pHelpSlave^.SlaveInfo.pPath = NIL then
              ClassState := -1;
              retcode := -2;
              return;
            end_if;

            // save hardwarepath
            _memcpy(ptr1:=pHelpSlave^.SlaveInfo.pPath, ptr2:=pDataHelp, cntr:=TmpPathLen);
            pDataHelp += TmpPathLen;

            // length of hardwarepath
            TmpPathLen := pDataHelp^$UINT; // save some time with this local variable
            pHelpSlave^.SlaveInfo.CompPathLen := TmpPathLen;
            pDataHelp += sizeof(UINT);

            // allocate memory for the module path
            pHelpSlave^.SlaveInfo.pCompPath$pVoid := To_StdLib.Malloc(size:=TmpPathLen);
            if pHelpSlave^.SlaveInfo.pCompPath = NIL then
              ClassState := -1;
              retcode := -2;
              return;
            end_if;

            // save compressed hardwarepath
            _memcpy(ptr1:=pHelpSlave^.SlaveInfo.pCompPath, ptr2:=pDataHelp, cntr:=TmpPathLen);
            pDataHelp += TmpPathLen;
          else
            ClassState := -1;
            retcode := -2;
            return;
          end_if;
        end_for;
      end_if;

      pHelpCfg^.pFirstFSoEConnection := NIL;

      // check if it's a FSoE Config
      if IsFSoEConfig then
        // number of connection details which follow now
        TempConnectionNo := pDataHelp^$UINT;
        pDataHelp += sizeof(UINT);

        // if we got connections
        if TempConnectionNo then
          for i := 0 to (TempConnectionNo-1) do
            if pHelpCfg^.pFirstFSoEConnection = NIL then
              pHelpCfg^.pFirstFSoEConnection$pVoid := To_StdLib.Malloc(size:=sizeof(t_FSoEConnectionDetails));
              pHelpConnection := pHelpCfg^.pFirstFSoEConnection;
            else
              pHelpConnection^.pNext$pvoid := To_StdLib.Malloc(size:=sizeof(t_FSoEConnectionDetails));
              pHelpConnection := pHelpConnection^.pNext;
            end_if;

            // if we succeeded to allocate memory
            if pHelpConnection then
              // initialize the pointers with NIL in case one of the mallocs fails
              pHelpConnection^.pSlavePath       := NIL;
              pHelpConnection^.pSlavePathComp   := NIL;
              pHelpConnection^.pNext            := NIL;
              pHelpConnection^.pNextSorted      := NIL;

              // connection ID
              pHelpConnection^.ConnectionID := pDataHelp^$UINT;
              pDataHelp += sizeof(UINT);

              // connection state (use our own state internally)
              pHelpConnection^.InternalConnectionState := FCS_RESET;
              pHelpConnection^.ConnectionState := pDataHelp^$t_FSoEConnectionState;

              pDataHelp += sizeof(USINT);

              // flags

              // Actually, type is 4 bytes in size but for compatibility reasons it is still used as 1 byte. As a result, bits 9-32 are currently not used.
              if bdFeatureEnable.FSoEFlags_4ByteSize then
                pHelpConnection^.Flags$t_FSoEFlags := pDataHelp^$t_FSoEFlags;
                pDataHelp += sizeof(t_FSoEFlags);
              else
                pHelpConnection^.Flags$USINT := pDataHelp^$USINT;
                pDataHelp += sizeof(USINT);
              end_if;

              // master safety number
              pHelpConnection^.OwnerSafetyNbr := pDataHelp^$HDINT;
              pDataHelp += sizeof(HDINT);

              // the feature is not available in older safety module classes, so we have to do this for compatibility reasons
              if bdFeatureEnable.TransmissionTimeInConfig then
                // transmission time in ms
                pHelpConnection^.TransmissionTime_ms := pDataHelp^$UINT;
                pDataHelp += sizeof(UINT);
              else
                pHelpConnection^.TransmissionTime_ms := 0;
              end_if;

              // offset where to read from master
              pHelpConnection^.MasterReadOffset := pDataHelp^$UINT;
              pDataHelp += sizeof(UINT);

              // size of data to read from master (and write to slave)
              pHelpConnection^.MasterReadSize := pDataHelp^$UINT;
              pDataHelp += sizeof(UINT);

              // offset where to write to master
              pHelpConnection^.MasterWriteOffset := pDataHelp^$UINT;
              pDataHelp += sizeof(UINT);

              // size of data to write to master (and read from slave)
              pHelpConnection^.MasterWriteSize := pDataHelp^$UINT;
              pDataHelp += sizeof(UINT);

              // slave address
              pHelpConnection^.SlaveAddress := pDataHelp^$UINT;
              pDataHelp += sizeof(UINT);

              // wait for slave addresses if any connection is not initialized
              if (pHelpConnection^.ConnectionState = FCS_NOT_INITIALIZED) & (pHelpConnection^.SlaveAddress = 0) then
                b_AllLocalSlaveAddressesValid := FALSE;
              end_if;

              // length of uncompressed slave hardwarepath
              TmpPathLen := pDataHelp^$UINT; // save some time with this local variable
              pHelpConnection^.SlavePathLen := TmpPathLen;
              pDataHelp += sizeof(UINT);

              if pHelpConnection^.Flags.IsMaster then
                // allocate memory for the module path
                pHelpConnection^.pSlavePath$pVoid := To_StdLib.Malloc(size:=TmpPathLen);
                if pHelpConnection^.pSlavePath = NIL then
                  ClassState := -1;
                  retcode := -2;
                  return;
                end_if;

                // save hardwarepath
                _memcpy(ptr1:=pHelpConnection^.pSlavePath, ptr2:=pDataHelp, cntr:=TmpPathLen);
                pDataHelp += TmpPathLen;
              end_if;

              // length of compressed slave hardwarepath
              TmpPathLen := pDataHelp^$UINT; // save some time with this local variable
              pHelpConnection^.SlavePathCompLen := TmpPathLen;
              pDataHelp += sizeof(UINT);

              if pHelpConnection^.Flags.IsMaster then
                // allocate memory for the module path
                pHelpConnection^.pSlavePathComp$pVoid := To_StdLib.Malloc(size:=TmpPathLen);
                if pHelpConnection^.pSlavePathComp = NIL then
                  ClassState := -1;
                  retcode := -2;
                  return;
                end_if;

                // save compressed hardwarepath
                _memcpy(ptr1:=pHelpConnection^.pSlavePathComp, ptr2:=pDataHelp, cntr:=TmpPathLen);
                pDataHelp += TmpPathLen;

                // if it's a udp connection, consider the transmission time
                if (pHelpConnection^.pSlavePathComp^ = INTERFACE_IP_MODE) & pHelpConnection^.TransmissionTime_ms then
                  if pHelpConnection^.TransmissionTime_ms < sUdpVars.LowestTransmissionTime_ms then
                    sUdpVars.LowestTransmissionTime_ms := pHelpConnection^.TransmissionTime_ms;
                  end_if;
                end_if;
              end_if;

              // offset where to read from master
              pHelpConnection^.SlaveReadOffset := pDataHelp^$UINT;
              pDataHelp += sizeof(UINT);

              // offset where to write to master
              pHelpConnection^.SlaveWriteOffset := pDataHelp^$UINT;
              pDataHelp += sizeof(UINT);

              // initialize log marker
              pHelpConnection^.bsLogError := 0;
            else
              ClassState := -1;
              retcode := -2;
              return;
            end_if;
          end_for;
        end_if;
      end_if;

      ConfigNo += 1;

      // check if the given size matches the memory structure
      if (pDataHelp$UDINT - pData$UDINT) <> Length then
        LogError("@ZZZZ (SafetyManager::AddConfiguration) Invalid configuration data given (length doesn't match memory structure)");
        retcode := -3;
        return;
      end_if;
    else
      ClassState := -1;
      retcode := -2;
      return;
    end_if;
  else
    // invalid configuration
    LogError("@ZZZZ (SafetyManager::AddConfiguration) Found invalid safety cpu configuration: Pointer or size wrong");
    retcode := -1;
  end_if;

END_FUNCTION

FUNCTION SafetyManager::FreeCfgLists
  VAR
    pHelpCfg        : ^t_CfgListElem;
    pHelpModule     : ^t_ModuleListElem;
    pHelpPdo        : ^t_PdoListElem;
    pHelpConnection : ^t_FSoEConnectionDetails;
  END_VAR

  while pConfigs do
    pHelpCfg := pConfigs;
    pConfigs := pConfigs^.pNext;

    // while we got module cfgs
    while pHelpCfg^.pFirstModuleCfg do
      pHelpModule := pHelpCfg^.pFirstModuleCfg;
      pHelpCfg^.pFirstModuleCfg := pHelpCfg^.pFirstModuleCfg^.pNext;

      if pHelpModule^.ModuleInfo.pDestCRCs then
        To_StdLib.Free(pHelpModule^.ModuleInfo.pDestCRCs);
      end_if;

      To_StdLib.Free(pHelpModule^.ModuleInfo.pPath);
      To_StdLib.Free(pHelpModule^.ModuleInfo.pCompPath);
      To_StdLib.Free(pHelpModule);
    end_while;

    // while we got pdo cfgs
    while pHelpCfg^.pFirstPdoCfg do
      pHelpPdo := pHelpCfg^.pFirstPdoCfg;
      pHelpCfg^.pFirstPdoCfg := pHelpCfg^.pFirstPdoCfg^.pNext;

      To_StdLib.Free(pHelpPdo^.PdoInfo.pSourcePath);
      To_StdLib.Free(pHelpPdo^.PdoInfo.pDestPath);
      To_StdLib.Free(pHelpPdo);
    end_while;

    // while we got connection infos
    while pHelpCfg^.pFirstFSoEConnection do
      pHelpConnection := pHelpCfg^.pFirstFSoEConnection;
      pHelpCfg^.pFirstFSoEConnection := pHelpCfg^.pFirstFSoEConnection^.pNext;

      if pHelpConnection^.pSlavePath then
        To_StdLib.Free(mptr:=pHelpConnection^.pSlavePath);
      end_if;

      if pHelpConnection^.pSlavePathComp then
        To_StdLib.Free(mptr:=pHelpConnection^.pSlavePathComp);
      end_if;

      To_StdLib.Free(mptr:=pHelpConnection);
    end_while;

    To_StdLib.Free(pHelpCfg);
  end_while;
  pSortedConnections := NIL; // may have contained a pointer within the config (to the connection with the lowest slave address)
  ConfigNo := 0;

END_FUNCTION

FUNCTION SafetyManager::AddOwnCPUsToList
  VAR
  	pHelpSafety : ^t_SafetyComponent;
  END_VAR

  // reset number of memorized safe cpu numbers
  SafeCPU_Nbr_No := 0;

  // check if any of the managing modules is not synchron
  if pFirstSafetyComponent then
    pHelpSafety := pFirstSafetyComponent;
    while pHelpSafety do
      // add all safety cpus to the parameters
      if IsCPUModule(pHelpSafety^.ModuleType) then
        if pHelpSafety^.SafetyNbr then
          aSafetyCPU_Nbr[SafeCPU_Nbr_No] := pHelpSafety^.SafetyNbr;
          SafeCPU_Nbr_No += 1;
        end_if;
      end_if;

      pHelpSafety := pHelpSafety^.pNext;
    end_while;
  end_if;

END_FUNCTION

FUNCTION SafetyManager::AllCPUConfigsArrived
	VAR_OUTPUT
		AllReady 	: BOOL;
	END_VAR
  VAR
    pHelpCfg : ^t_CfgListElem;
    i : UDINT;
    Found : BOOL;
  END_VAR

  // check if there are any CPUs
  if SafeCPU_Nbr_No then
    // if we have already all configurations (according to the number) check if they are correct
    if ConfigNo = SafeCPU_Nbr_No then

      // normally we should be fine now
      AllReady := TRUE;

      // check all safety numbers stored
      for i := 0 to SafeCPU_Nbr_No-1 do

        Found := FALSE;

        // search all configurations
        pHelpCfg := pConfigs;
        while pHelpCfg do
          // if we found a match => stop searching for this one
          if pHelpCfg^.SafetyNbr = aSafetyCPU_Nbr[i] then
            Found := TRUE;
            exit;
          end_if;
          pHelpCfg := pHelpCfg^.pNext;
        end_while;

        // if this configuration hasn't been found, we may have a problem
        if Found = FALSE then
          AllReady := FALSE;
          LogError("@ZZZZ (SafetyManager::AllCPUConfigsArrived) Invalid CPU configuration found!");
          return;
        end_if;
      end_for;
    else
      AllReady := FALSE;

      if ConfigNo > SafeCPU_Nbr_No then
        LogError("@ZZZZ (SafetyManager::AllCPUConfigsArrived) ERROR! More configs available than safety CPUs");
      end_if;
    end_if;
  else
    AllReady := TRUE;
    LogError("@ZZZZ (SafetyManager::AllCPUConfigsArrived) No Safety CPU found in the system!");
  end_if;

END_FUNCTION

FUNCTION SafetyManager::AddLocalCPUCfg
	VAR_INPUT
		Length 	: UINT;
		pData 	: ^void;
		IsFSoECfg 	: BOOL;(* := FALSE *)
	END_VAR
  VAR
  	pHelpLocalCfg   : ^t_LocalCfgListElem;
    EditOldCfg      : BOOL;
  END_VAR

  LastCfgReceiveTime := ops.tAbsolute;

  // if the a module wants to add the config which is already added => overwrite the old config
  EditOldCfg := FALSE;

  if pFirstLocalCPUCfg = NIL then
    pFirstLocalCPUCfg$pVoid := To_StdLib.Malloc(size:=sizeof(t_LocalCfgListElem));
    pHelpLocalCfg := pFirstLocalCPUCfg;
  else
    pHelpLocalCfg := pFirstLocalCPUCfg;

    if pHelpLocalCfg^.SafetyNbr = pData^$HDINT then
      EditOldCfg := TRUE;
    else
      while pHelpLocalCfg^.pNext <> NIL do
        pHelpLocalCfg := pHelpLocalCfg^.pNext;
        if pHelpLocalCfg^.SafetyNbr = pData^$HDINT then
          EditOldCfg := TRUE;
          exit;
        end_if;
      end_while;
      if EditOldCfg = FALSE then
        pHelpLocalCfg^.pNext$pVoid := To_StdLib.Malloc(size:=sizeof(t_LocalCfgListElem));

        pHelpLocalCfg := pHelpLocalCfg^.pNext;
      end_if;
    end_if;
  end_if;

  if pHelpLocalCfg <> NIL then
    pHelpLocalCfg^.SafetyNbr          := pData^$HDINT;
    pHelpLocalCfg^.ConfigSize         := Length;
    pHelpLocalCfg^.pConfig            := pData;  // memory can be accessed always (never freed)
    pHelpLocalCfg^.ConfigSent2Master  := FALSE;
    pHelpLocalCfg^.IsFSoECfg          := IsFSoECfg;

    if IsFSoECfg then
      sUdpVars.UdpInit.FSoEAvailable := TRUE;
    end_if;

    // only if we created a new element (incrementing has to be done last becuase of thread safety: bg increments the value and cyclic uses the list)
    if EditOldCfg = FALSE then
      pHelpLocalCfg^.pNext := NIL;
      LocalCPUCfgNo += 1;

      // new cpu config => reinitalize everything
      ReinitEverything();
    end_if;
  else
    ClassState := -1;
    LogError("@ZZZZ (SafetyManager::AddLocalCPUCfg) Failed to allocate Memory for the local CPU Configuration");
  end_if;

END_FUNCTION

FUNCTION SafetyManager::SendLocalCfgsToMaster
  VAR
  	pHelpLocalCfg : ^t_LocalCfgListElem;
    i : UDINT;
  END_VAR

  if LocalCPUCfgNo then
    pHelpLocalCfg := pFirstLocalCPUCfg;

    for i := 0 to (LocalCPUCfgNo-1) do
      if pHelpLocalCfg^.ConfigSize then
        // if we're the master, we keep the configuration of this cpu and share the essentials later (when we got all configurations) with all other domains (distribute the mapping)
        if AddConfiguration(pHelpLocalCfg^.ConfigSize, pHelpLocalCfg^.pConfig, pHelpLocalCfg^.IsFSoECfg) <> 0 then
          LogError("@ZZZZ (SafetyManager::SendLocalCfgsToMaster) Failed to add a safety cpu configuration to the local config-memory");
        end_if;
      end_if;

      pHelpLocalCfg := pHelpLocalCfg^.pNext;
    end_for;
  end_if;

END_FUNCTION

FUNCTION SafetyManager::BroadCastActPDO
  VAR
		MyPara 	  : CmdStruct;
    PdoMemSize : UINT;
    pPdoMem    : ^USINT;
    pHelp      : ^USINT;
    TmpPathLen : UINT;
    SourceDest : t_SourceDest;
    SafetyNbr           : HDINT;
  END_VAR

  // put pdo (marked by pActualSendPDO) into linear memory, find out who needs it and broadcast it

(*
    Memory structure:
      1 Byte: Number of Domains involved
      x Byte: 1 Byte for every involved Domain number
      1 Byte: Number of Domains in source path
      x Byte: 1 Byte for every domain in source path
      1 Byte: Number of Domains in destination path
      x Byte: 1 Byte for every domain in destination path
      1 Byte: ID of this PDO (starting at 0)
      1 Byte: Length of PDO
      1 Byte: Is it an interface frame
      4 Byte: Interface CRC
      2 Byte: Length of source hardware path
      x Byte (depending on length in the 2 byte before): Hardwarepath of source
      2 Byte: Length of destination hardware path
      x Byte (depending on length in the 2 byte before): Hardwarepath of destination
*)

  // if the pointer is NIL or it's an interface frame broadcast, don't distribute it, there are virtual PDOs to be distributed instead of the broadcasts (if necessary)
  if (pActualSendPDO = NIL) | pActualSendPDO^.PdoInfo.Info.IFBroadCast then
    return;
  end_if;

  // add up the sizes and allocate the memory
  PdoMemSize := sizeof(USINT) +                           // 1 byte number of domains involved
                1 +                                       // 1 byte for every involved domain
                sizeof(USINT) +                           // 1 byte number of domains in source path
                1 +                                       // 1 byte for every domain in source path
                sizeof(USINT) +                           // 1 byte number of domains in destination path
                1 +                                       // 1 byte for every domain in destination path
                sizeof(USINT) +                           // 1 byte ID of this PDO (starting at 0)
                sizeof(USINT) +                           // 1 byte length of PDO
                sizeof(t_PdoCfgInfo) +                    // 1 byte pdo info (is it interface frame or optional...)
                sizeof(HDINT) +                           // 4 byte interface CRC
                sizeof(UINT) +                            // 2 byte length of source hardware path
                pActualSendPDO^.PdoInfo.SourcePathLen +   // x byte source hardware path
                sizeof(UINT) +                            // 2 byte length of destination hardware path
                pActualSendPDO^.PdoInfo.DestPathLen;      // x byte destination hardware path

  if ud_SizeTempMemCy >= PdoMemSize then
    pPdoMem := pTempMemCy$^USINT;
  else
    LogError("@ZZZZ (SafetyManager::BroadCastActPDO) Temporary memory for cyclic task is too small!");
    LogValue("AvaliableMem: {0} / NeededMem: {1}", Value:=ud_SizeTempMemCy, Value2:=PdoMemSize);
    ClassState := -1;
    return;
  end_if;

  if pPdoMem then
    pHelp := pPdoMem;

    // number of domains involved
    pHelp^$USINT := 1;
    pHelp += sizeof(USINT);

    // domain number of this ack
    pHelp^$USINT := 0;
    pHelp += 1;

    // number of domains in source path
    pHelp^$USINT := 1;
    pHelp += sizeof(USINT);

    // domain numbers of source domains
    pHelp^$USINT := 0;
    pHelp += 1;

    // number of domains in dest path
    pHelp^$USINT := 1;
    pHelp += sizeof(USINT);

    // domain numbers of dest domains
    pHelp^$USINT := 0;
    pHelp += 1;

    pHelp^$USINT := pActualSendPDO^.PdoInfo.PDO_ID;
    pHelp += sizeof(USINT);

    pHelp^$USINT := pActualSendPDO^.PdoInfo.PdoLen;
    pHelp += sizeof(USINT);

    pHelp^$t_PdoCfgInfo := pActualSendPDO^.PdoInfo.Info;
    pHelp += sizeof(t_PdoCfgInfo);

    pHelp^$HDINT := pActualSendPDO^.PdoInfo.InterfaceCRC;
    pHelp += sizeof(HDINT);

    TmpPathLen := pActualSendPDO^.PdoInfo.SourcePathLen; // save some time with this local variable
    pHelp^$UINT := TmpPathLen;
    pHelp += sizeof(UINT);

    _memcpy(ptr1:=pHelp, ptr2:=pActualSendPDO^.PdoInfo.pSourcePath, cntr:=TmpPathLen);
    pHelp += TmpPathLen;

    TmpPathLen := pActualSendPDO^.PdoInfo.DestPathLen;
    pHelp^$UINT := TmpPathLen;
    pHelp += sizeof(UINT);

    _memcpy(ptr1:=pHelp, ptr2:=pActualSendPDO^.PdoInfo.pDestPath, cntr:=TmpPathLen);

    MyPara.uiCmd := CMD_SM_PDO_MAPPING_BROADCAST;
    MyPara.aPara[0] := PdoMemSize; // length of parameters
    MyPara.aPara[1] := pPdoMem$DINT;

    // check out if we have to work with this, and if so save the PDO info's
    if IsAffectedByPDO(#MyPara, #SourceDest, #SafetyNbr) then

    end_if;
  else
    ClassState := -1;
    LogError("@ZZZZ (SafetyManager::BroadCastActPDO) Failed to allocate memory for the currently broadcasting PDO Info");
  end_if;

END_FUNCTION

FUNCTION SafetyManager::IsAffectedByPDO
	VAR_INPUT
		pPara 	: ^CmdStruct;
		pSourceDest 	: ^t_SourceDest;
		pSafetyNbr 	: ^HDINT;
	END_VAR
	VAR_OUTPUT
		IsAffected 	: BOOL;
	END_VAR
  VAR
  	pHelp                 :^USINT;
    pFirstDomainAffected  : ^USINT;
    DomainsInside         : USINT;
    SourcePathLen         : UINT;
    pSourcePath           : ^USINT;
    DestPathLen           : UINT;
    pDestPath             : ^USINT;
    pHelpManaging         : ^t_ManagingComponent;
    pHelpSafety           : ^t_SafetyComponent;
    pSourceSafety         : ^t_SafetyComponent;
    pDestSafety           : ^t_SafetyComponent;
		MyPara 	              : CmdStruct;
		MyResult	            : results;
    PDO_ID                : USINT;
    Length                : USINT;
    SourceDomain          : USINT;
    DestDomain            : USINT;
    SourceDomainNo        : USINT;
    DestDomainNo          : USINT;
    aSourceDomains        : ARRAY [0..99] OF USINT;
    aDestDomains          : ARRAY [0..99] OF USINT;
    IsInterfaceFrame      : BOOL;
    InterfaceCRC          : HDINT;
    CopyCmdIndex          : INT;
    pPDOElement           : ^t_PDOElement;
    pRecyclePDO           : ^t_PDOElement;
    TempLen               : USINT;
    TempOffset            : UDINT;
    PDOInfo               : t_PdoCfgInfo;
  END_VAR

  IsAffected := FALSE;

  pSourceDest^ := SourceDest_None;
  pSafetyNbr^ := 0;

  // check the parameters
  pFirstDomainAffected := (pPara^.aPara[1])$^USINT;
  pHelp  := pFirstDomainAffected;

  DomainsInside := pHelp^$USINT;
  pHelp += sizeof(USINT);

  if DomainsInside then
    // skip the domain number
    pHelp += sizeof(USINT);

    IsAffected := TRUE;

(*
    Memory structure:
      1 Byte: Number of Domains involved
      x Byte: 1 Byte for every involved Domain number
      1 Byte: Number of Domains in source path
      x Byte: 1 Byte for every domain in source path
      1 Byte: Number of Domains in destination path
      x Byte: 1 Byte for every domain in destination path
      1 Byte: ID of this PDO (starting at 0)
      1 Byte: Length of PDO
      1 Byte: PDO Info (Is it an interface frame, or optional...)
      4 Byte: Interface CRC
      2 Byte: Length of source hardware path
      x Byte (depending on length in the 2 byte before): Hardwarepath of source
      2 Byte: Length of destination hardware path
      x Byte (depending on length in the 2 byte before): Hardwarepath of destination
*)

    if IsAffected then
      // pHelp is now pointing to the Number of Domains in source path

      _memset(dest:=#aSourceDomains[0], usByte:=16#FF, cntr:=sizeof(aSourceDomains));
      _memset(dest:=#aDestDomains[0], usByte:=16#FF, cntr:=sizeof(aDestDomains));

      SourceDomainNo := pHelp^;
      pHelp += sizeof(USINT);

      _memcpy(ptr1:=#aSourceDomains[0], ptr2:=pHelp, cntr:=SourceDomainNo);
      pHelp += SourceDomainNo;

      DestDomainNo := pHelp^;
      pHelp += sizeof(USINT);

      _memcpy(ptr1:=#aDestDomains[0], ptr2:=pHelp, cntr:=DestDomainNo);
      pHelp += DestDomainNo;

      PDO_ID := pHelp^;
      pHelp += sizeof(USINT);

      Length := pHelp^;
      pHelp += sizeof(USINT);

      PDOInfo := pHelp^;
      IsInterfaceFrame := PDOInfo.IsInterfacePDO;
      pHelp += sizeof(t_PdoCfgInfo);

      InterfaceCRC := pHelp^$HDINT;
      pHelp += sizeof(HDINT);

      SourcePathLen := pHelp^$UINT;
      pHelp += sizeof(UINT);
      pSourcePath := pHelp;
      pHelp += SourcePathLen;
      DestPathLen := pHelp^$UINT;
      pHelp += sizeof(UINT);
      pDestPath := pHelp;

      SourceDomain := aSourceDomains[SourceDomainNo-1];
      DestDomain   := aDestDomains[DestDomainNo-1];

      pSourceSafety := NIL;
      pDestSafety   := NIL;

      // if we're the source or destination domain and there is a safety component in this system, check if it's the source or destination for this PDO
      if pFirstSafetyComponent then
        // check for source or dest module
        pHelpSafety := pFirstSafetyComponent;
        while pHelpSafety & ((pSourceSafety = NIL) | (pDestSafety = NIL)) do
          // we compare the last x byte (where x is the length of the local path including the domain)
          if (pSourceSafety = NIL) then
            // if the length matches it's in the same domain, otherwise the local search path must be shorter and there must be a domain escape sequence in the long path
            if pHelpSafety^.pPath & ((pSourcePath^ = pHelpSafety^.pPath^) | ((pSourcePath^ > pHelpSafety^.pPath^) & ((pSourcePath + 1 + pSourcePath^ - pHelpSafety^.pPath^)^ = HWT_ESCAPE_DOMAIN))) &
               (To_StdLib.MemCmp(pHelpSafety^.pPath + 1, pSourcePath + 2 + pSourcePath^ - pHelpSafety^.pPath^, pHelpSafety^.pPath^) = 0) then

              pSourceSafety := pHelpSafety;
            end_if;
          end_if;

          if (pDestSafety = NIL) then
            // if the length matches it's in the same domain, otherwise the local search path must be shorter and there must be a domain escape sequence in the long path
            if pHelpSafety^.pPath & ((pDestPath^ = pHelpSafety^.pPath^) | ((pDestPath^ > pHelpSafety^.pPath^) & ((pDestPath + 1 + pDestPath^ - pHelpSafety^.pPath^)^ = HWT_ESCAPE_DOMAIN))) &
               (To_StdLib.MemCmp(pHelpSafety^.pPath + 1, pDestPath + 2 + pDestPath^ - pHelpSafety^.pPath^, pHelpSafety^.pPath^) = 0) then

              pDestSafety := pHelpSafety;
              AddTimeSyncElement(pManaging:=NIL, pSafety:=pHelpSafety, IsInterfaceDomain := FALSE);
            end_if;
          end_if;

          pHelpSafety := pHelpSafety^.pNext;
        end_while;
      end_if;

      // use the pointer to the array element to save time
      pPDOElement := #aPDOElements[PDOElementNo];

      // here we have to check what to do with the PDO:
      // is the actual domain the source or the destination domain? or maybe both?
      if pSourceSafety & pDestSafety then
        pSourceDest^ := SourceDest_IsSourceAndDest;

        // only possible for interface frames
        if IsInterfaceFrame then
          // we have to tell the source, that there's a receiver for the PDO (also get the addresses)
          MyPara.uiCmd := CMD_SM_ADD_OUTPUT_PDO;
          MyPara.aPara[0] := 1;  // mark as interface frame PDO

          pSourceSafety^.pThis^.NewInst(#MyPara, #MyResult);

          // use a PDO element for automated removal of the input pdo in case of a new config
          pPDOElement^.PDO_ID                   := PDO_ID;
          pPDOElement^.Length                   := Length;
          pPDOElement^.ThisDomainsRole          := SourceDest_IsDest;
          pPDOElement^.SourceInfo.pPDOMem       := MyResult.aData[0]$^USINT;
          pPDOElement^.SourceInfo.pPDOMemDPRAM  := MyResult.aData[4]$^USINT;
          pPDOElement^.SourceInfo.SafetyNbr     := pSourceSafety^.SafetyNbr;
          pPDOElement^.DestInfo.SafetyNbr       := pDestSafety^.SafetyNbr;
          pPDOElement^.pSafety                  := pDestSafety;
          pPDOElement^.SourceInfo.HandlePDODPRAM:= MyResult.aData[8]$UDINT;   // Needed for Payload Support
          pPDOElement^.SourceInfo.OffsetPDODPRAM:= MyResult.aData[12]$UDINT;  // Needed for Payload Support
          PDOElementNo += 1;

          // then tell the destination about the PDO
          MyPara.uiCmd := CMD_SM_ADD_INPUT_PDO;
          MyPara.aPara[0] := pPDOElement^.SourceInfo.pPDOMem$DINT;  // we got the pointer to the local mem and the pointer to the DPRAM from the call of the source module
          MyPara.aPara[1] := pPDOElement^.SourceInfo.pPDOMemDPRAM$DINT;
          MyPara.aPara[2] := pSourceSafety^.SafetyNbr$DINT;
          MyPara.aPara[3] := Length;
          MyPara.aPara[4] := pActualSendPDO^.PdoInfo.Info.IsOptional; // only possible because this kind of PDOs is only available on Domain 0
          MyPara.aPara[5] := pPDOElement^.SourceInfo.HandlePDODPRAM$DINT; // Needed for Payload Support
          MyPara.aPara[6] := pPDOElement^.SourceInfo.OffsetPDODPRAM$DINT; // Needed for Payload Support
          MyPara.aPara[7] := 0;// target offset (not necessary here)
          MyPara.aPara[8] := SM_IF_VALIDITY_MARK$DINT;
          MyPara.aPara[9] := TRUE;

          pDestSafety^.pThis^.NewInst(#MyPara, #MyResult);
        else
          LogError("@ZZZZ (SafetyManager::IsAffectedByPDO) Error in PDO distribution: No InterfaceFrame but Source and Destination in this domain!");
        end_if;
      elsif pSourceSafety & (pDestSafety = NIL) then
        pSourceDest^ := SourceDest_IsSource;

        // get safety number of the source
        MyPara.uiCmd := CMD_SM_GET_SAFETY_NUMBER;
        MyPara.aPara[0] := pSafetyNbr$DINT;
        pSourceSafety^.pThis^.NewInst(#MyPara, #MyResult);

        pPDOElement^.PDO_ID                 := PDO_ID;
        pPDOElement^.Length                 := Length;
        pPDOElement^.ThisDomainsRole        := SourceDest_IsSource;

        pPDOElement^.SourceInfo.SafetyNbr   := pSafetyNbr^;
        pPDOElement^.SourceInfo.DomainNr    := SourceDomain;
        pPDOElement^.SourceInfo.PathLen     := SourcePathLen;
        pPDOElement^.SourceInfo.pPath$pVoid := To_StdLib.Malloc(size:= SourcePathLen);
        if pPDOElement^.SourceInfo.pPath then
          _memcpy(ptr1:=pPDOElement^.SourceInfo.pPath, ptr2:=pSourcePath, cntr:=SourcePathLen);
        else
          LogError("@ZZZZ (SafetyManager::IsAffectedByPDO) Failed to allocate memory for PDO path info");
          ClassState := -1;
          return;
        end_if;

        pPDOElement^.DestInfo.SafetyNbr     := 0;
        pPDOElement^.DestInfo.DomainNr      := DestDomain;
        pPDOElement^.DestInfo.PathLen       := DestPathLen;
        pPDOElement^.DestInfo.pPath$pVoid   := To_StdLib.Malloc(size:= DestPathLen);
        if pPDOElement^.DestInfo.pPath then
          _memcpy(ptr1:=pPDOElement^.DestInfo.pPath, ptr2:=pDestPath, cntr:=DestPathLen);
        else
          LogError("@ZZZZ (SafetyManager::IsAffectedByPDO) Failed to allocate memory for PDO path info");
          ClassState := -1;
          return;
        end_if;

        pPDOElement^.pSafety              := pSourceSafety;

        // initialize with invalid;
        CopyCmdIndex := -1;

        // if we're the master, we may also route interfaceframes
        if IsInterfaceFrame then
          // search for the destination of this PDO
          pHelpManaging := pFirstManagingInterfaceComponent;
          while pHelpManaging do
            if (To_StdLib.MemCmp(pHelpManaging^.pModulePath, pDestPath, DestPathLen) = 0) then
              exit;
            else
              pHelpManaging := pHelpManaging^.pNext;
            end_if;
          end_while;

          pPDOElement^.pManagingDest := pHelpManaging;
        end_if;

        if pPDOElement^.pManagingDest then

          // if the module is marked as optional and the PDO is not optional => the module is also not optional
          if pPDOElement^.pManagingDest^.InfoBits.IsOptional & (PDOInfo.IsOptional = FALSE) then
            pPDOElement^.pManagingDest^.InfoBits.IsOptional  := FALSE;
          end_if;

          // check if we can recycle the memory of another DO (if this data is already transferred to this managing module
          pRecyclePDO := CheckPDORecycle(SourceDest_IsDest, pPDOElement);

          // only if there is enough space or we already have a memory
          if pRecyclePDO | ((pPDOElement^.pManagingDest^.PDOWriteMemUsed + pPDOElement^.Length) <= pPDOElement^.pManagingDest^.PDOWriteMemAvailable) then

            // if we can't use the copy command
            if b_SafetyOnLocalCDIAS then
              // remember the pointer to the memory to copy it manually in rt postscan method
              if pRecyclePDO then
                // this PDO is already in the memory of the managing node, we don't have to copy it again
                pPDOElement^.DestInfo.pPDOMem := NIL;//pRecyclePDO^.DestInfo.pPDOMem;
              else
                pPDOElement^.DestInfo.pPDOMem := pPDOElement^.pManagingDest^.pPDOWriteSpace + pPDOElement^.pManagingDest^.PDOWriteMemUsed;
              end_if;
            else
              if pRecyclePDO then
                // this PDO is already in the memory of the managing node, we don't have to copy it again
                pPDOElement^.DestInfo.pPDOMemDPRAM := NIL;//pRecyclePDO^.DestInfo.pPDOMemDPRAM;
              else
                pPDOElement^.DestInfo.pPDOMemDPRAM := pPDOElement^.pManagingDest^.pPDOWriteSpaceDPRAM + pPDOElement^.pManagingDest^.PDOWriteMemUsed;
              end_if;

              CopyCmdIndex := GetNewMovDO();
              if CopyCmdIndex < 0 then
                if pRecyclePDO then
                  // this PDO is already in the memory of the managing node, we don't have to copy it again
                  pPDOElement^.DestInfo.pPDOMem := NIL;//pRecyclePDO^.DestInfo.pPDOMem;
                else
                  pPDOElement^.DestInfo.pPDOMem := pPDOElement^.pManagingDest^.pPDOWriteSpace + pPDOElement^.pManagingDest^.PDOWriteMemUsed;
                end_if;
                LogError("@ZZZZ (SafetyManager::IsAffectedByPDO) Failed to install copy command => PDO is beeing copied in RT");
              else
                aCopyCmds[CopyCmdIndex].pSettings^.ud_AddressDest := pPDOElement^.DestInfo.pPDOMemDPRAM$UDINT;
                aCopyCmds[CopyCmdIndex].pSettings^.ui_ByteCnt     := pPDOElement^.Length;
              end_if;
            end_if;

            // if we need new memory, tell the managing module
            if pRecyclePDO = NIL then
              pPDOElement^.pManagingDest^.PDOWriteMemUsed += pPDOElement^.Length;

              MyPara.uiCmd := CMD_SM_PDO_MEM_USAGE_WR;
              MyPara.aPara[0] := pPDOElement^.pManagingDest^.PDOWriteMemUsed$DINT;
              pPDOElement^.pManagingDest^.pThis^.NewInst(#MyPara, #MyResult);
            end_if;

            if IsInterfaceFrame then
              MyPara.uiCmd := CMD_SM_ADD_OUTPUT_PDO;
              MyPara.aPara[0] := 1;  // mark as interface frame PDO
              pSourceSafety^.pThis^.NewInst(#MyPara, #MyResult);

              pPDOElement^.SourceInfo.pPDOMem       := MyResult.aData[0]$^USINT;
              pPDOElement^.SourceInfo.pPDOMemDPRAM  := MyResult.aData[4]$^USINT;
              pPDOElement^.SourceInfo.HandlePDODPRAM:= MyResult.aData[8]$UDINT;   // Needed for Payload Support
              pPDOElement^.SourceInfo.OffsetPDODPRAM:= MyResult.aData[12]$UDINT;  // Needed for Payload Support
            end_if;
          else
            // we add the memory anyway to show the user how much he would need
            pPDOElement^.pManagingDest^.PDOWriteMemUsed += pPDOElement^.Length;

            MyPara.uiCmd := CMD_SM_PDO_MEM_USAGE_WR;
            MyPara.aPara[0] := pPDOElement^.pManagingDest^.PDOWriteMemUsed$DINT;
            pPDOElement^.pManagingDest^.pThis^.NewInst(#MyPara, #MyResult);

            LogError("@ZZZZ (SafetyManager::IsAffectedByPDO) Not enough write memory to map all PDOs");
            return;
          end_if;
        else
          LogError("@ZZZZ (SafetyManager::IsAffectedByPDO) Couldn't find destination managing module for PDO");
          return;
        end_if;

        pPDOElement^.CopyCmdIndex := CopyCmdIndex;

        PDOElementNo += 1;
      elsif pDestSafety & (pSourceSafety = NIL) then
        pSourceDest^ := SourceDest_IsDest;

        // get safety number of the destination
        MyPara.uiCmd := CMD_SM_GET_SAFETY_NUMBER;
        MyPara.aPara[0] := pSafetyNbr$DINT;
        pDestSafety^.pThis^.NewInst(#MyPara, #MyResult);

        pPDOElement^.PDO_ID                 := PDO_ID;
        pPDOElement^.Length                 := Length;
        pPDOElement^.ThisDomainsRole        := SourceDest_IsDest;

        pPDOElement^.SourceInfo.SafetyNbr   := 0;
        pPDOElement^.SourceInfo.DomainNr    := SourceDomain;
        pPDOElement^.SourceInfo.PathLen     := SourcePathLen;
        pPDOElement^.SourceInfo.pPath$pVoid := To_StdLib.Malloc(size:= SourcePathLen);
        if pPDOElement^.SourceInfo.pPath then
          _memcpy(ptr1:=pPDOElement^.SourceInfo.pPath, ptr2:=pSourcePath, cntr:=SourcePathLen);
        else
          LogError("@ZZZZ (SafetyManager::IsAffectedByPDO) Failed to allocate memory for PDO path info");
          ClassState := -1;
          return;
        end_if;

        pPDOElement^.DestInfo.SafetyNbr     := pSafetyNbr^;
        pPDOElement^.DestInfo.DomainNr      := DestDomain;
        pPDOElement^.DestInfo.PathLen       := DestPathLen;
        pPDOElement^.DestInfo.pPath$pVoid   := To_StdLib.Malloc(size:= DestPathLen);
        if pPDOElement^.DestInfo.pPath then
          _memcpy(ptr1:=pPDOElement^.DestInfo.pPath, ptr2:=pDestPath, cntr:=DestPathLen);
        else
          LogError("@ZZZZ (SafetyManager::IsAffectedByPDO) Failed to allocate memory for PDO path info");
          ClassState := -1;
          return;
        end_if;

        pPDOElement^.pSafety              := pDestSafety;

        // if we're the master, we may also route interfaceframes
        if IsInterfaceFrame then

          // search for the source of this PDO
          pHelpManaging := pFirstManagingInterfaceComponent;
          while pHelpManaging do
            if (To_StdLib.MemCmp(pHelpManaging^.pModulePath, pSourcePath, SourcePathLen) = 0) then
              exit;
            else
              pHelpManaging := pHelpManaging^.pNext;
            end_if;
          end_while;

          pPDOElement^.pManagingSource := pHelpManaging;
        end_if;

        if pPDOElement^.pManagingSource then

          // if the module is marked as optional and the PDO is not optional => the module is also not optional
          if pPDOElement^.pManagingSource^.InfoBits.IsOptional & (PDOInfo.IsOptional = FALSE) then
            pPDOElement^.pManagingSource^.InfoBits.IsOptional  := FALSE;
          end_if;

          // check if we can recycle the memory of another DO (if this data is already transferred to this managing module
          pRecyclePDO := CheckPDORecycle(SourceDest_IsSource, pPDOElement);

          // only if there is enough space or we already have a memory
          if pRecyclePDO | ((pPDOElement^.pManagingSource^.PDOReadMemUsed + pPDOElement^.Length) <= pPDOElement^.pManagingSource^.PDOReadMemAvailable) then
            if IsInterfaceFrame then
              pPDOElement^.SourceInfo.SafetyNbr   := (GetIFInfoByCRC(InterfaceCRC, #TempOffset, #TempLen))$HDINT;
              if TempLen = Length then
                // get the place in the memory of the source managing module
                pPDOElement^.SourceInfo.pPDOMem       := pPDOElement^.pManagingSource^.pPDOReadSpace + TempOffset;
                pPDOElement^.SourceInfo.pPDOMemDPRAM  := pPDOElement^.pManagingSource^.pPDOReadSpaceDPRAM + TempOffset;

                pPDOElement^.SourceInfo.HandlePDODPRAM := pPDOElement^.pManagingSource^.ud_HandlePDOReadSpaceDPRAM;
                pPDOElement^.SourceInfo.OffsetPDODPRAM := TempOffset;

                // if we need new memory, tell the managing module
                if (TempOffset + Length) > pPDOElement^.pManagingSource^.PDOReadMemUsed then
                  pPDOElement^.pManagingSource^.PDOReadMemUsed := TempOffset + Length;

                  MyPara.uiCmd := CMD_SM_PDO_MEM_USAGE_RD;
                  MyPara.aPara[0] := pPDOElement^.pManagingSource^.PDOReadMemUsed$DINT;
                  pPDOElement^.pManagingSource^.pThis^.NewInst(#MyPara, #MyResult);
                end_if;

                MyPara.uiCmd := CMD_SM_ADD_INPUT_PDO;
                MyPara.aPara[0] := pPDOElement^.SourceInfo.pPDOMem$DINT;
                MyPara.aPara[1] := pPDOElement^.SourceInfo.pPDOMemDPRAM$DINT;
                MyPara.aPara[2] := pPDOElement^.SourceInfo.SafetyNbr$DINT;
                MyPara.aPara[3] := Length;
                MyPara.aPara[4] := PDOInfo.IsOptional;
                MyPara.aPara[5] := pPDOElement^.SourceInfo.HandlePDODPRAM$DINT; // Needed for Payload Support
                MyPara.aPara[6] := pPDOElement^.SourceInfo.OffsetPDODPRAM$DINT; // Needed for Payload Support
                MyPara.aPara[7] := 0;// target offset (not necessary here)
                MyPara.aPara[8] := SM_IF_VALIDITY_MARK$DINT;
                MyPara.aPara[9] := TRUE;

                pDestSafety^.pThis^.NewInst(#MyPara, #MyResult);
              else
                LogError("@ZZZZ (SafetyManager::IsAffectedByPDO) Length of interface frames doesn't match the local configuration");
              end_if;

            else
              if pRecyclePDO then
                pPDOElement^.SourceInfo.pPDOMem       := pRecyclePDO^.SourceInfo.pPDOMem;
                pPDOElement^.SourceInfo.pPDOMemDPRAM  := pRecyclePDO^.SourceInfo.pPDOMemDPRAM;
              else
                pPDOElement^.SourceInfo.pPDOMem       := pPDOElement^.pManagingSource^.pPDOReadSpace + pPDOElement^.pManagingSource^.PDOReadMemUsed;
                pPDOElement^.SourceInfo.pPDOMemDPRAM  := pPDOElement^.pManagingSource^.pPDOReadSpaceDPRAM + pPDOElement^.pManagingSource^.PDOReadMemUsed;

                // if we need new memory, tell the managing module
                pPDOElement^.pManagingSource^.PDOReadMemUsed += pPDOElement^.Length;

                MyPara.uiCmd := CMD_SM_PDO_MEM_USAGE_RD;
                MyPara.aPara[0] := pPDOElement^.pManagingSource^.PDOReadMemUsed$DINT;
                pPDOElement^.pManagingSource^.pThis^.NewInst(#MyPara, #MyResult);
              end_if;
            end_if;
          else
            // we add the memory anyway to show the user how much he would need
            pPDOElement^.pManagingSource^.PDOReadMemUsed += pPDOElement^.Length;

            MyPara.uiCmd := CMD_SM_PDO_MEM_USAGE_RD;
            MyPara.aPara[0] := pPDOElement^.pManagingSource^.PDOReadMemUsed$DINT;
            pPDOElement^.pManagingSource^.pThis^.NewInst(#MyPara, #MyResult);

            LogError("@ZZZZ (SafetyManager::IsAffectedByPDO) Not enough read memory to map all PDOs");
            return;
          end_if;
        else

          LogError("@ZZZZ (SafetyManager::IsAffectedByPDO) Couldn't find source managing module for PDO");
          return;
        end_if;

        PDOElementNo += 1;
      else
        pSourceDest^ := SourceDest_IsForwarder;

        // if source and destination are not in this domain, is it a bifurcation or a linear forwarding?
        pPDOElement^.PDO_ID                 := PDO_ID;
        pPDOElement^.Length                 := Length;
        pPDOElement^.ThisDomainsRole        := SourceDest_IsForwarder;

        pPDOElement^.SourceInfo.DomainNr    := SourceDomain;
        pPDOElement^.SourceInfo.PathLen     := SourcePathLen;
        pPDOElement^.SourceInfo.pPath$pVoid := To_StdLib.Malloc(size:= SourcePathLen);
        if pPDOElement^.SourceInfo.pPath then
          _memcpy(ptr1:=pPDOElement^.SourceInfo.pPath, ptr2:=pSourcePath, cntr:=SourcePathLen);
        else
          LogError("@ZZZZ (SafetyManager::IsAffectedByPDO) Failed to allocate memory for PDO path info");
          ClassState := -1;
          return;
        end_if;

        pPDOElement^.DestInfo.DomainNr      := DestDomain;
        pPDOElement^.DestInfo.PathLen       := DestPathLen;
        pPDOElement^.DestInfo.pPath$pVoid   := To_StdLib.Malloc(size:= DestPathLen);
        if pPDOElement^.DestInfo.pPath then
          _memcpy(ptr1:=pPDOElement^.DestInfo.pPath, ptr2:=pDestPath, cntr:=DestPathLen);
        else
          LogError("@ZZZZ (SafetyManager::IsAffectedByPDO) Failed to allocate memory for PDO path info");
          ClassState := -1;
          return;
        end_if;

        // initialize with invalid;
        CopyCmdIndex := -1;

        // if we're the master, we may also route interfaceframes
        if IsInterfaceFrame then

          // search for the source of this PDO
          pHelpManaging := pFirstManagingInterfaceComponent;
          while pHelpManaging do
            if (To_StdLib.MemCmp(pHelpManaging^.pModulePath, pSourcePath, SourcePathLen) = 0) then
              exit;
            else
              pHelpManaging := pHelpManaging^.pNext;
            end_if;
          end_while;

          pPDOElement^.pManagingSource := pHelpManaging;
        end_if;

        if pPDOElement^.pManagingSource then

          // if the module is marked as optional and the PDO is not optional => the module is also not optional
          if pPDOElement^.pManagingSource^.InfoBits.IsOptional & (PDOInfo.IsOptional = FALSE) then
            pPDOElement^.pManagingSource^.InfoBits.IsOptional  := FALSE;
          end_if;

          // check if we can recycle the memory of another DO (if this data is already transferred to this managing module
          pRecyclePDO := CheckPDORecycle(SourceDest_IsSource, pPDOElement);

          if pRecyclePDO | ((pPDOElement^.pManagingSource^.PDOReadMemUsed + pPDOElement^.Length) <= pPDOElement^.pManagingSource^.PDOReadMemAvailable) then
            if pRecyclePDO then
              pPDOElement^.SourceInfo.pPDOMem       := pRecyclePDO^.SourceInfo.pPDOMem;
              pPDOElement^.SourceInfo.pPDOMemDPRAM  := pRecyclePDO^.SourceInfo.pPDOMemDPRAM;
            else
              pPDOElement^.SourceInfo.pPDOMem       := pPDOElement^.pManagingSource^.pPDOReadSpace + pPDOElement^.pManagingSource^.PDOReadMemUsed;
              pPDOElement^.SourceInfo.pPDOMemDPRAM  := pPDOElement^.pManagingSource^.pPDOReadSpaceDPRAM + pPDOElement^.pManagingSource^.PDOReadMemUsed;
              pPDOElement^.pManagingSource^.PDOReadMemUsed += pPDOElement^.Length;

              MyPara.uiCmd := CMD_SM_PDO_MEM_USAGE_RD;
              MyPara.aPara[0] := pPDOElement^.pManagingSource^.PDOReadMemUsed$DINT;
              pPDOElement^.pManagingSource^.pThis^.NewInst(#MyPara, #MyResult);
            end_if;
          else
            // we add the memory anyway to show the user how much he would need
            pPDOElement^.pManagingSource^.PDOReadMemUsed += pPDOElement^.Length;

            MyPara.uiCmd := CMD_SM_PDO_MEM_USAGE_RD;
            MyPara.aPara[0] := pPDOElement^.pManagingSource^.PDOReadMemUsed$DINT;
            pPDOElement^.pManagingSource^.pThis^.NewInst(#MyPara, #MyResult);

            LogError("@ZZZZ (SafetyManager::IsAffectedByPDO) Not enough read memory to map all PDOs");
            return;
          end_if;
        else
          LogError("@ZZZZ (SafetyManager::IsAffectedByPDO) Couldn't find source managing module for PDO");
          return;
        end_if;

        // if we're the master, we may also route interfaceframes
        if IsInterfaceFrame then
          // search for the destination of this PDO
          pHelpManaging := pFirstManagingInterfaceComponent;
          while pHelpManaging do
            if (To_StdLib.MemCmp(pHelpManaging^.pModulePath, pDestPath, DestPathLen) = 0) then
              exit;
            else
              pHelpManaging := pHelpManaging^.pNext;
            end_if;
          end_while;

          pPDOElement^.pManagingDest := pHelpManaging;
        end_if;

        if pPDOElement^.pManagingDest then

          // if the module is marked as optional and the PDO is not optional => the module is also not optional
          if pPDOElement^.pManagingDest^.InfoBits.IsOptional & (PDOInfo.IsOptional = FALSE) then
            pPDOElement^.pManagingDest^.InfoBits.IsOptional  := FALSE;
          end_if;

          if pPDOElement^.pManagingDest = pPDOElement^.pManagingSource then
            LogError("@ZZZZ (SafetyManager::IsAffectedByPDO) In PDO Forwarding a domain can't be the source and the destination!");
          end_if;

          // check if we can recycle the memory of another DO (if this data is already transferred to this managing module
          pRecyclePDO := CheckPDORecycle(SourceDest_IsDest, pPDOElement);

          if pRecyclePDO | ((pPDOElement^.pManagingDest^.PDOWriteMemUsed + pPDOElement^.Length) <= pPDOElement^.pManagingDest^.PDOWriteMemAvailable) then

            // if we can't use the copy command
            if b_SafetyOnLocalCDIAS then
              // remember the pointer to the memory to copy it manually in rt postscan method
              if pRecyclePDO then
                // this PDO is already in the memory of the managing node, we don't have to copy it again
                pPDOElement^.DestInfo.pPDOMem := NIL;//pRecyclePDO^.SourceInfo.pPDOMem;
              else
                pPDOElement^.DestInfo.pPDOMem := pPDOElement^.pManagingDest^.pPDOWriteSpace + pPDOElement^.pManagingDest^.PDOWriteMemUsed;
              end_if;
            else
              if pRecyclePDO then
                // this PDO is already in the memory of the managing node, we don't have to copy it again
                pPDOElement^.DestInfo.pPDOMemDPRAM := NIL;//pRecyclePDO^.DestInfo.pPDOMemDPRAM;
              else
                pPDOElement^.DestInfo.pPDOMemDPRAM := pPDOElement^.pManagingDest^.pPDOWriteSpaceDPRAM + pPDOElement^.pManagingDest^.PDOWriteMemUsed;
              end_if;

              CopyCmdIndex := GetNewMovDO();
              if CopyCmdIndex < 0 then
                pPDOElement^.DestInfo.pPDOMem := pPDOElement^.pManagingDest^.pPDOWriteSpace + pPDOElement^.pManagingDest^.PDOWriteMemUsed;
                LogError("@ZZZZ (SafetyManager::IsAffectedByPDO) Failed to install copy command => PDO is beeing copied in RT");
              else
                aCopyCmds[CopyCmdIndex].pSettings^.ud_AddressDest := pPDOElement^.DestInfo.pPDOMemDPRAM$UDINT;
                aCopyCmds[CopyCmdIndex].pSettings^.ui_ByteCnt     := pPDOElement^.Length;
              end_if;
            end_if;

            // if we need new memory, tell the managing module
            if pRecyclePDO = NIL then
              pPDOElement^.pManagingDest^.PDOWriteMemUsed += pPDOElement^.Length;

              MyPara.uiCmd := CMD_SM_PDO_MEM_USAGE_WR;
              MyPara.aPara[0] := pPDOElement^.pManagingDest^.PDOWriteMemUsed$DINT;
              pPDOElement^.pManagingDest^.pThis^.NewInst(#MyPara, #MyResult);
            end_if;
          else
            // we add the memory anyway to show the user how much he would need
            pPDOElement^.pManagingDest^.PDOWriteMemUsed += pPDOElement^.Length;

            MyPara.uiCmd := CMD_SM_PDO_MEM_USAGE_WR;
            MyPara.aPara[0] := pPDOElement^.pManagingDest^.PDOWriteMemUsed$DINT;
            pPDOElement^.pManagingDest^.pThis^.NewInst(#MyPara, #MyResult);

            LogError("@ZZZZ (SafetyManager::IsAffectedByPDO) Not enough write memory to map all PDOs");
            return;
          end_if;
        else
          LogError("@ZZZZ (SafetyManager::IsAffectedByPDO) Couldn't find destination managing module for PDO");
          return;
        end_if;

        pPDOElement^.CopyCmdIndex := CopyCmdIndex;

        PDOElementNo += 1;
      end_if;

    end_if;
  end_if;

END_FUNCTION

FUNCTION SafetyManager::GetDestManagingOfDO
	VAR_INPUT
		pDO 	: ^SafetyCDIAS_Base::SDOHeader;
	END_VAR
	VAR_OUTPUT
		pDestManaging 	: ^t_ManagingComponent;
	END_VAR
	VAR
		pHelpManaging 	: ^t_ManagingComponent;
    i : UDINT;
	END_VAR

  pDestManaging := NIL;

  // maybe it's one of the interface domains
  pHelpManaging := pFirstManagingInterfaceComponent;
  while pHelpManaging do
    if pHelpManaging^.ModuleNo then
      for i := 0 to (pHelpManaging^.ModuleNo-1) do
        if pHelpManaging^.ModuleInfo[i].SafetyNbr = pDO^.DstAdr then
          pDestManaging := pHelpManaging;
          return;
        end_if;
      end_for;
    end_if;

    pHelpManaging := pHelpManaging^.pNext;
  end_while;

END_FUNCTION

FUNCTION SafetyManager::GetDestSafetyOfDO
	VAR_INPUT
		pDO 	: ^SafetyCDIAS_Base::SDOHeader;
	END_VAR
	VAR_OUTPUT
		pDestSafety 	: ^t_SafetyComponent;
	END_VAR
	VAR
		pHelpSafety 	: ^t_SafetyComponent;
	END_VAR

  pDestSafety := NIL;

  // check if it's a SDO addressed via safety number
  if (pDO^.StdHeader.Typ AND SSDO_MASK_TYPE) = FRM_TYPECODE_SSDO_MOD_TP then
    // we can't find it via Topology path
    LogError("@ZZZZ (SafetyManager::GetDestSafetyOfDO) Misdirected SDO via Topology path. Addressee can't be found here");
    return;
  end_if;

  pHelpSafety := pFirstSafetyComponent;
  while pHelpSafety do
    if pHelpSafety^.SafetyNbr = pDO^.DstAdr then
      pDestSafety := pHelpSafety;
      return;
    end_if;

    pHelpSafety := pHelpSafety^.pNext;
  end_while;

END_FUNCTION

FUNCTION VIRTUAL GLOBAL SafetyManager::RtWork
	VAR_INPUT
		EAX 	: UDINT;
	END_VAR
	VAR_OUTPUT
		state (EAX) 	: UDINT;
	END_VAR
  VAR
  	i                 : UDINT;
    pPDOElement       : ^t_PDOElement;
    pFSoEElement      : ^t_FSoECopyCmd;
    AllCopyCmdsReady  : BOOL;
  END_VAR

  if EAX = CALL_OPTION_RT_PRESCAN then
    // prescan

//=================================================================================================
#ifdef VM_CLASS_TIME_MEASUREMENT
	StartTimeMeasurement(VARANTIME_RT);
#endif
//=================================================================================================

    // copy commands for udp connections (receiving via udp)
    if sUdpVars.ReceiveCopyCmdNo then
      // we may have some udp send data, so we better protect the copy mechanism
      UdpReceiveData.SectionStart();

      pFSoEElement := #sUdpVars.aReceiveCopyCmds[0];
      for i := 1 to sUdpVars.ReceiveCopyCmdNo do
        _memcpy(ptr1:=pFSoEElement^.pDest, ptr2:=pFSoEElement^.pSource, cntr:=pFSoEElement^.Size);
        pFSoEElement += sizeof(t_FSoECopyCmd);
      end_for;

      UdpReceiveData.SectionStop();
    end_if;

    case InitSSW of
//**********************************************************************************************************************************************************
      _Wait4CopyCmdStart:
        // start all used copy commands
        AllCopyCmdsReady := TRUE;
        if CopyCmdsUsed then
          for i := 0 to (CopyCmdsUsed-1) do
            if aCopyCmds[i].b_Ready4Action then
              aCopyCmds[i].pHandle^.ucCtrlStat := VARAN_DO_CONT_RUN;
            else
              AllCopyCmdsReady := FALSE;
              bd_LogRtMessagesInCy.UnkownCopySource := TRUE;
            end_if;
          end_for;
        end_if;

        if AllCopyCmdsReady then
          InitSSW := _FinishInitialisation;
        end_if;

//**********************************************************************************************************************************************************
      _InitFinished:
        // if we're master or we're actually time synchronizing
        if b_NewSyncMode & b_CheckTimeSyncTimeout then
          if (ops.tAbsolute - TimeSyncTimeStamp) > TIMESYNC_TIMEOUT then
            // increment timeout counter => message is shown in cyclic after x consecutive
            SyncTimeoutCounter += 1;
            b_CheckTimeSyncTimeout := FALSE; // => show Trace Message only once per error
            // restart the synchronisation (maybe the other domain has been disconnected)
            b_StartTimeSync := TRUE;
          end_if;
        end_if;

//**********************************************************************************************************************************************************
    end_case;

    // marker is set in cyclic priority (except on timeout), but time synchronisation has to be done in rt priority => start it from here
    if b_StartTimeSync then
      b_StartTimeSync := FALSE;

      StartTimeSync();
    end_if;

//=================================================================================================
#ifdef VM_CLASS_TIME_MEASUREMENT
	StopTimeMeasurement(VARANTIME_RT);
#endif
//=================================================================================================

  else
    // postscan

//=================================================================================================
#ifdef VM_CLASS_TIME_MEASUREMENT
	StartTimeMeasurement(VARANTIME_RTPOSTSCAN);
#endif
//=================================================================================================

    // copy data from our memory to the memory of the next domain
    if PDOElementNo then
      pPDOElement := #aPDOElements[0];
      for i := 1 to PDOElementNo do
        if (pPDOElement^.ThisDomainsRole = SourceDest_IsSource) |
           (pPDOElement^.ThisDomainsRole = SourceDest_IsForwarder) then
          if pPDOElement^.DestInfo.pPDOMem & pPDOElement^.SourceInfo.pPDOMem & pPDOElement^.Length then
            _memcpy(ptr1:=pPDOElement^.DestInfo.pPDOMem, ptr2:=pPDOElement^.SourceInfo.pPDOMem, cntr:=pPDOElement^.Length);
          end_if;
        end_if;
        pPDOElement += sizeof(t_PDOElement);
      end_for;
    elsif FSoECopyCmdNo then
      pFSoEElement := #aFSoECopyCmds[0];
      for i := 1 to FSoECopyCmdNo do
        _memcpy(ptr1:=pFSoEElement^.pDest, ptr2:=pFSoEElement^.pSource, cntr:=pFSoEElement^.Size);
        pFSoEElement += sizeof(t_FSoECopyCmd);
      end_for;
    end_if;

    // copy commands for udp connections (sending via udp)
    if sUdpVars.SendCopyCmdNo then
      // we may have some udp send data, so we better protect the copy mechanism
      UdpSendData.SectionStart();

      pFSoEElement := #sUdpVars.aSendCopyCmds[0];
      for i := 1 to sUdpVars.SendCopyCmdNo do
        _memcpy(ptr1:=pFSoEElement^.pDest, ptr2:=pFSoEElement^.pSource, cntr:=pFSoEElement^.Size);
        pFSoEElement += sizeof(t_FSoECopyCmd);
      end_for;

      UdpSendData.SectionStop();
    end_if;

//=================================================================================================
#ifdef VM_CLASS_TIME_MEASUREMENT
	StopTimeMeasurement(VARANTIME_RTPOSTSCAN);
#endif
//=================================================================================================

  end_if;

#ifdef SAFETY_DEBUG_LOGGING_ACTIVATED
  if InitSSW <> OldInitSSW then
#ifdef SAFETY_DEBUG_TRACING_ACTIVATED
    LogValue("@ZZZZ (SafetyManager::RtWork) InitSSW changed from {0} to {1}", Value:=OldInitSSW, Value2:=InitSSW);
#endif
    LogBuf[ActLogIndex].NewState := InitSSW;
    LogBuf[ActLogIndex].OldState := OldInitSSW;
    LogBuf[ActLogIndex].Command := 0;
    LogBuf[ActLogIndex].TimeSinceLastLog_us := OS_READMICROSEC();
    LogBuf[ActLogIndex].TimeSinceLastLog_us -= TimeStampLastLog_us;
    TimeStampLastLog_us := OS_READMICROSEC();
    if ActLogIndex = (LogBufferSize - 1) then
      ActLogIndex := 0;
    else
      ActLogIndex += 1;
    end_if;
  end_if;
  OldInitSSW := InitSSW;
#endif

	state := READY;

END_FUNCTION

FUNCTION SafetyManager::CheckTopSDO
	VAR_INPUT
		pPara 	: ^CmdStruct;
	END_VAR
  VAR
    pDO 	            : ^SafetyCDIAS_Base::SDOHeader;
    pCompDestPath     : ^USINT;
    pHelpConfig       : ^t_CfgListElem;
    pHelpSlave        : ^t_SlaveListElem;
    pHelpModule       : ^t_ModuleListElem;
    pHelpPdo          : ^t_PdoListElem;
    pHelpManaging     : ^t_ManagingComponent;
    pHelpSafety       : ^t_SafetyComponent;
    pHelpConnection   : ^t_FSoEConnectionDetails;
    MyPara            : CmdStruct;
    MyResult          : results;
    pTempMem          : ^USINT;
    pHelp             : ^USINT;
    TmpLen            : UINT;
    DomainChangeFound : BOOL;
    i                 : UDINT;
    DestDomain        : USINT;
    InterfaceCRC      : HDINT;
    TargetSafetyNbr   : HDINT;
    pActConnection    : ^t_UdpConnection;
  END_VAR

  // get a pointer to the compressed destination path
  pDO := (pPara^.aPara[1])$^SafetyCDIAS_Base::SDOHeader;
  pCompDestPath := (#pDO^.DstAdr)$^USINT;

  // if we have interfaceframes, check them first
  if pFirstManagingInterfaceComponent & (pCompDestPath^ = INTERFACE_CRC_MODE) then
    // after the mode byte we find the interface CRC
    InterfaceCRC := ((pCompDestPath + 1)$^HDINT)^;
